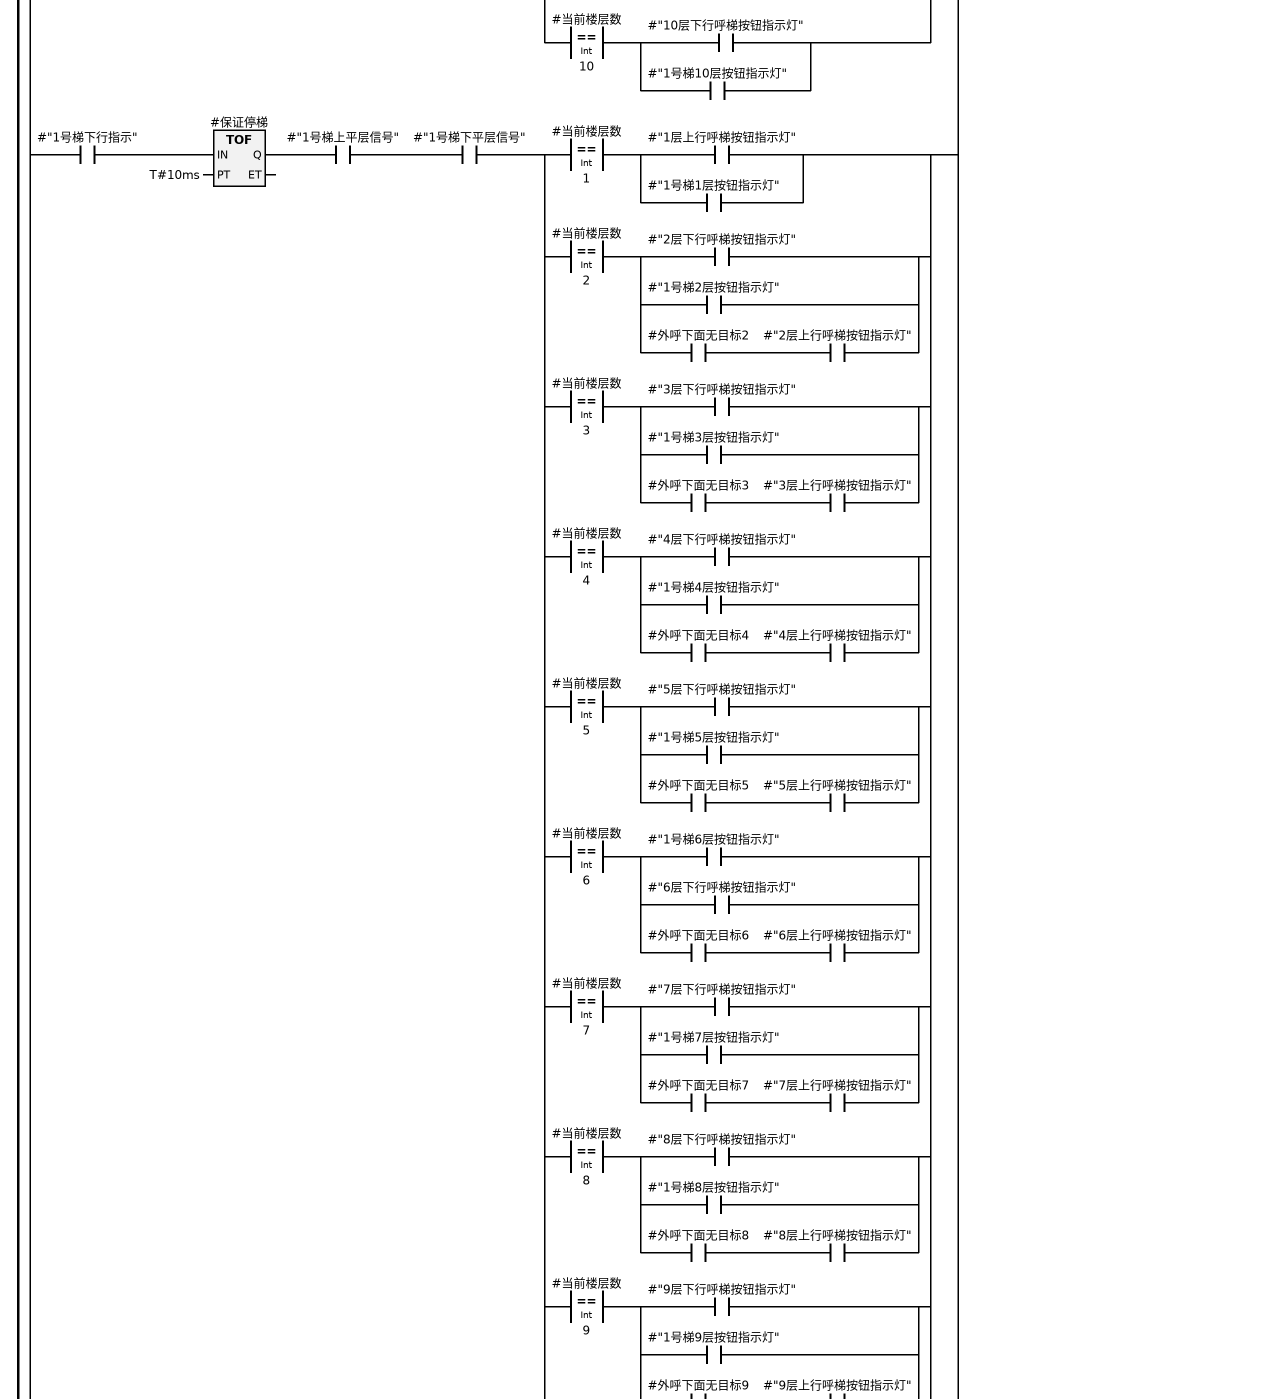
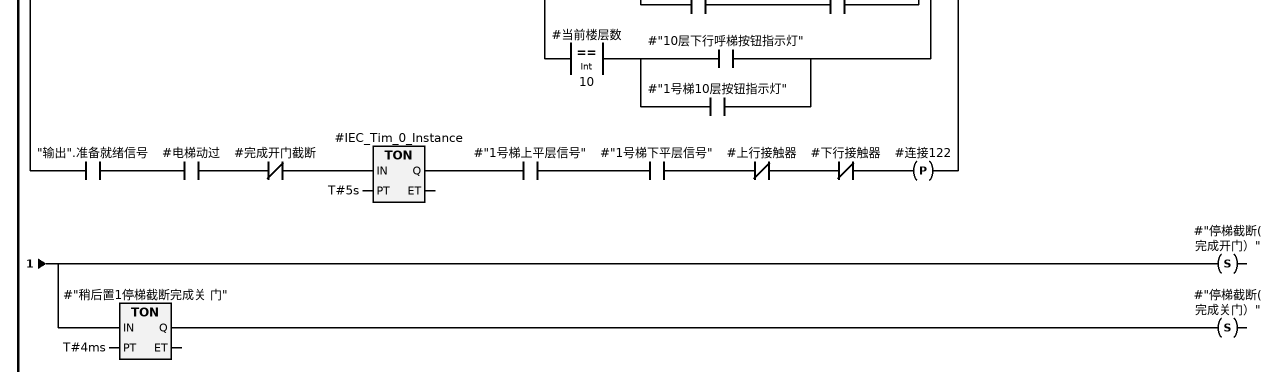
   #保证停梯上(IN := #"1号梯上行指示", PT := T#10ms);   // TOF
   #保证停梯(IN := #"1号梯下行指示", PT := T#10ms);   // TOF
   #IEC_Tim_0_Instance(IN := "输出".准备就绪信号 AND #电梯动过 AND NOT #完成开门截断, PT := T#5s);   // TON
   #_w1 := #IEC_Tim_0_Instance.Q AND #"1号梯上平层信号" AND #"1号梯下平层信号" AND NOT #上行接触器 AND NOT #下行接触器;
   #_w2 := #_w1 AND NOT #连接122;   // rising edge
   #连接122 := #_w1;
   #_w3 := ((#保证停梯上.Q AND #"1号梯上平层信号" AND #"1号梯下平层信号" AND (((#当前楼层数 = 1) AND (#"1层上行呼梯按钮指示灯" OR #"1号梯1层按钮指示灯")) OR ((#当前楼层数 = 2) AND (#"2层上行呼梯按钮指示灯" OR #"1号梯2层按钮指示灯" OR (#外呼上面无目标2 AND #"2层下行呼梯按钮指示灯"))) OR ((#当前楼层数 = 3) AND (#"3层上行呼梯按钮指示灯" OR #"1号梯3层按钮指示灯" OR (#外呼上面无目标3 AND #"3层下行呼梯按钮指示灯"))) OR ((#当前楼层数 = 4) AND (#"4层上行呼梯按钮指示灯" OR #"1号梯4层按钮指示灯" OR (#外呼上面无目标4 AND #"4层下行呼梯按钮指示灯"))) OR ((#当前楼层数 = 5) AND (#"5层上行呼梯按钮指示灯" OR #"1号梯5层按钮指示灯" OR (#外呼上面无目标5 AND #"5层下行呼梯按钮指示灯"))) OR ((#当前楼层数 = 6) AND (#"6层上行呼梯按钮指示灯" OR #"1号梯6层按钮指示灯" OR (#外呼上面无目标6 AND #"6层下行呼梯按钮指示灯"))) OR ((#当前楼层数 = 7) AND (#"7层上行呼梯按钮指示灯" OR #"1号梯7层按钮指示灯" OR (#外呼上面无目标7 AND #"7层下行呼梯按钮指示灯"))) OR ((#当前楼层数 = 8) AND (#"8层上行呼梯按钮指示灯" OR #"1号梯8层按钮指示灯" OR (#外呼上面无目标8 AND #"8层下行呼梯按钮指示灯"))) OR ((#当前楼层数 = 9) AND (#"9层上行呼梯按钮指示灯" OR #"1号梯9层按钮指示灯" OR (#外呼上面无目标9 AND #"9层下行呼梯按钮指示灯"))) OR ((#当前楼层数 = 10) AND (#"10层下行呼梯按钮指示灯" OR #"1号梯10层按钮指示灯")))) OR (#保证停梯.Q AND #"1号梯上平层信号" AND #"1号梯下平层信号" AND (((#当前楼层数 = 1) AND (#"1层上行呼梯按钮指示灯" OR #"1号梯1层按钮指示灯")) OR ((#当前楼层数 = 2) AND (#"2层下行呼梯按钮指示灯" OR #"1号梯2层按钮指示灯" OR (#外呼下面无目标2 AND #"2层上行呼梯按钮指示灯"))) OR ((#当前楼层数 = 3) AND (#"3层下行呼梯按钮指示灯" OR #"1号梯3层按钮指示灯" OR (#外呼下面无目标3 AND #"3层上行呼梯按钮指示灯"))) OR ((#当前楼层数 = 4) AND (#"4层下行呼梯按钮指示灯" OR #"1号梯4层按钮指示灯" OR (#外呼下面无目标4 AND #"4层上行呼梯按钮指示灯"))) OR ((#当前楼层数 = 5) AND (#"5层下行呼梯按钮指示灯" OR #"1号梯5层按钮指示灯" OR (#外呼下面无目标5 AND #"5层上行呼梯按钮指示灯"))) OR ((#当前楼层数 = 6) AND (#"1号梯6层按钮指示灯" OR #"6层下行呼梯按钮指示灯" OR (#外呼下面无目标6 AND #"6层上行呼梯按钮指示灯"))) OR ((#当前楼层数 = 7) AND (#"7层下行呼梯按钮指示灯" OR #"1号梯7层按钮指示灯" OR (#外呼下面无目标7 AND #"7层上行呼梯按钮指示灯"))) OR ((#当前楼层数 = 8) AND (#"8层下行呼梯按钮指示灯" OR #"1号梯8层按钮指示灯" OR (#外呼下面无目标8 AND #"8层上行呼梯按钮指示灯"))) OR ((#当前楼层数 = 9) AND (#"9层下行呼梯按钮指示灯" OR #"1号梯9层按钮指示灯" OR (#外呼下面无目标9 AND #"9层上行呼梯按钮指示灯"))) OR ((#当前楼层数 = 10) AND (#"10层下行呼梯按钮指示灯" OR #"1号梯10层按钮指示灯")))) OR #_w2) AND NOT #"1号梯检修信号" AND NOT #开门次数达到上限;
   IF #_w3 THEN #"停梯截断(完成开门）" := TRUE; END_IF;
   #"稍后置1停梯截断完成关 门"(IN := #_w3, PT := T#4ms);   // TON
   IF #"稍后置1停梯截断完成关 门".Q THEN #"停梯截断(完成关门）" := TRUE; END_IF;
END_REGION

REGION Network 2: 停梯后自主 开门
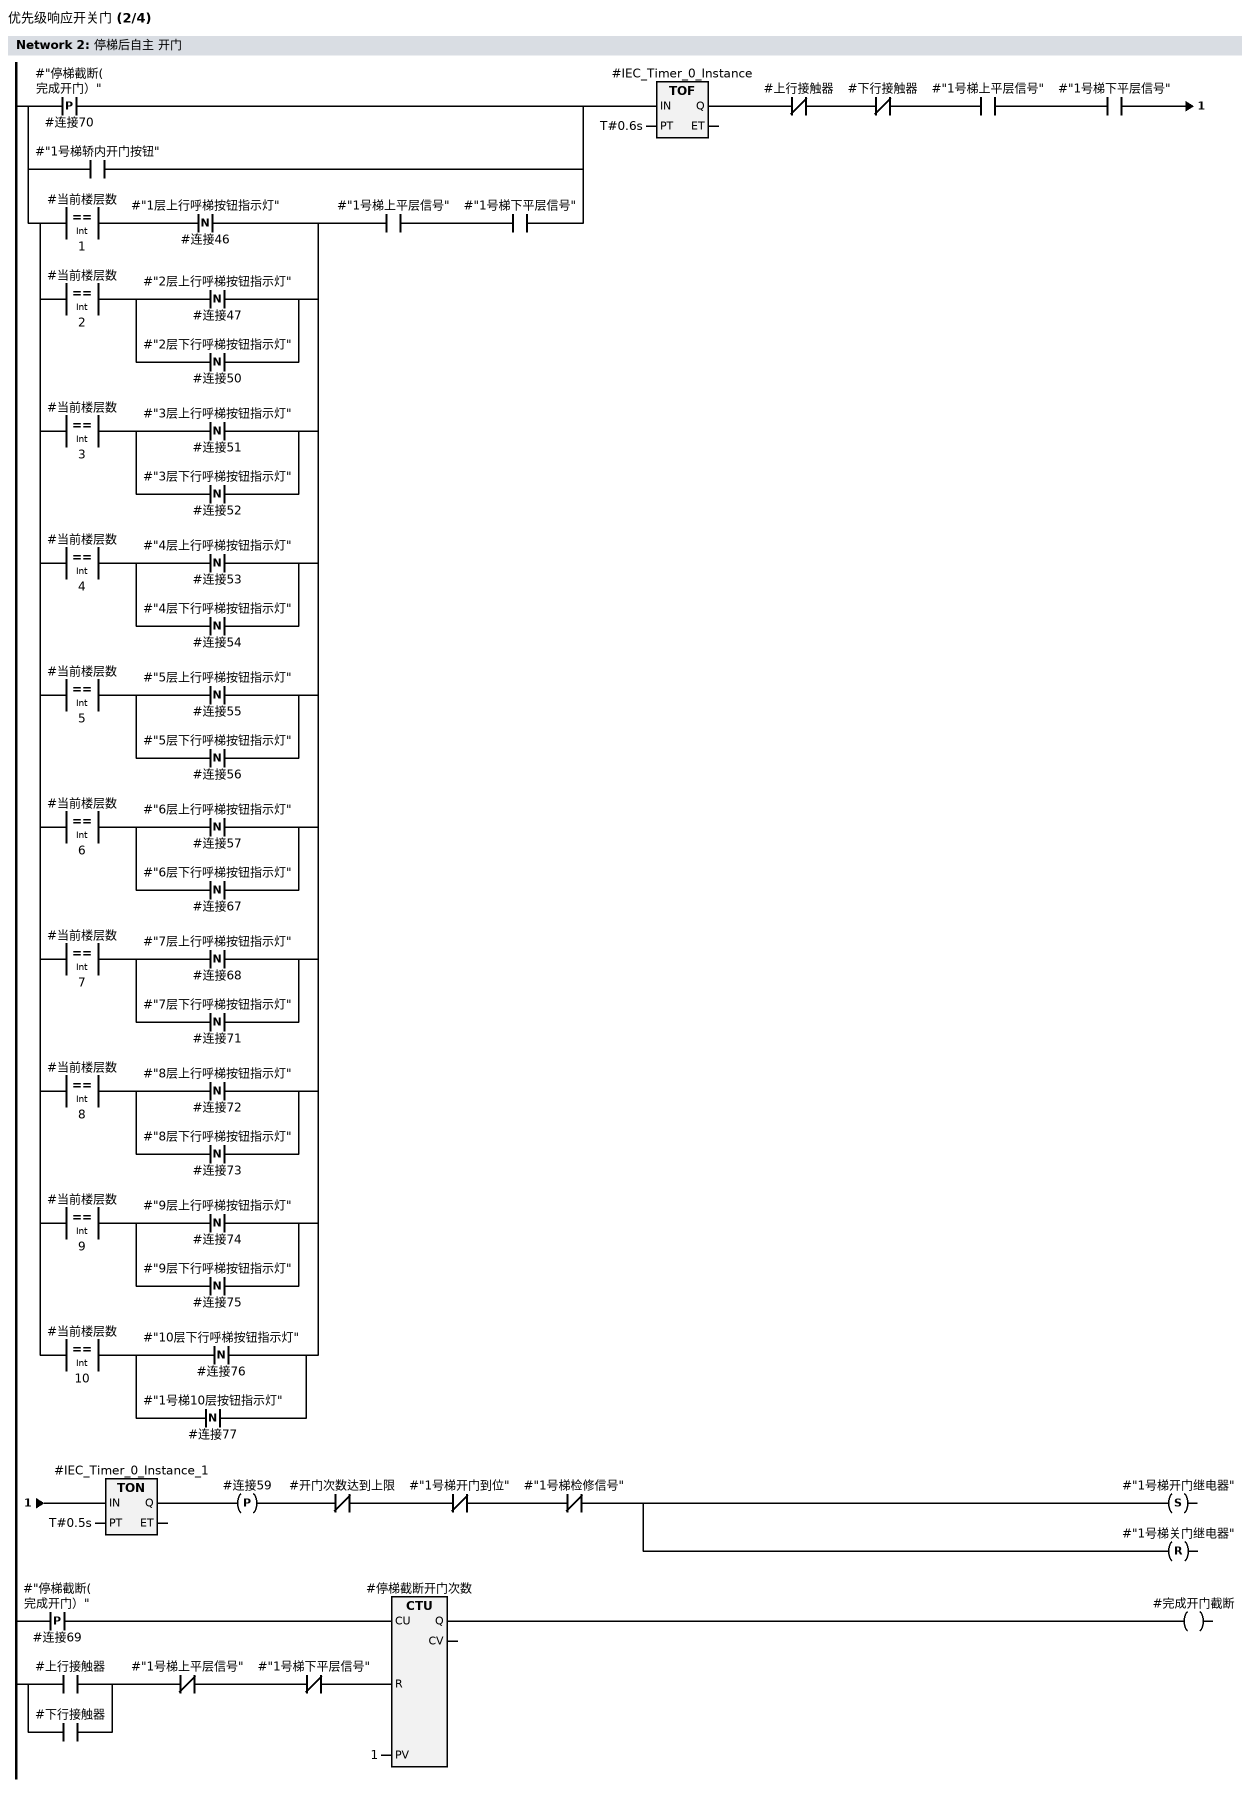
   #_w1 := #"停梯截断(完成开门）" AND NOT #连接70;   // rising edge of #"停梯截断(完成开门）"
   #连接70 := #"停梯截断(完成开门）";
   #_w2 := (#当前楼层数 = 1) AND NOT #"1层上行呼梯按钮指示灯" AND #连接46;   // falling edge of #"1层上行呼梯按钮指示灯"
   #连接46 := #"1层上行呼梯按钮指示灯";
   #_w3 := (#当前楼层数 = 2) AND NOT #"2层上行呼梯按钮指示灯" AND #连接47;   // falling edge of #"2层上行呼梯按钮指示灯"
   #连接47 := #"2层上行呼梯按钮指示灯";
   #_w4 := (#当前楼层数 = 2) AND NOT #"2层下行呼梯按钮指示灯" AND #连接50;   // falling edge of #"2层下行呼梯按钮指示灯"
   #连接50 := #"2层下行呼梯按钮指示灯";
   #_w5 := (#当前楼层数 = 3) AND NOT #"3层上行呼梯按钮指示灯" AND #连接51;   // falling edge of #"3层上行呼梯按钮指示灯"
   #连接51 := #"3层上行呼梯按钮指示灯";
   #_w6 := (#当前楼层数 = 3) AND NOT #"3层下行呼梯按钮指示灯" AND #连接52;   // falling edge of #"3层下行呼梯按钮指示灯"
   #连接52 := #"3层下行呼梯按钮指示灯";
   #_w7 := (#当前楼层数 = 4) AND NOT #"4层上行呼梯按钮指示灯" AND #连接53;   // falling edge of #"4层上行呼梯按钮指示灯"
   #连接53 := #"4层上行呼梯按钮指示灯";
   #_w8 := (#当前楼层数 = 4) AND NOT #"4层下行呼梯按钮指示灯" AND #连接54;   // falling edge of #"4层下行呼梯按钮指示灯"
   #连接54 := #"4层下行呼梯按钮指示灯";
   #_w9 := (#当前楼层数 = 5) AND NOT #"5层上行呼梯按钮指示灯" AND #连接55;   // falling edge of #"5层上行呼梯按钮指示灯"
   #连接55 := #"5层上行呼梯按钮指示灯";
   #_w10 := (#当前楼层数 = 5) AND NOT #"5层下行呼梯按钮指示灯" AND #连接56;   // falling edge of #"5层下行呼梯按钮指示灯"
   #连接56 := #"5层下行呼梯按钮指示灯";
   #_w11 := (#当前楼层数 = 6) AND NOT #"6层上行呼梯按钮指示灯" AND #连接57;   // falling edge of #"6层上行呼梯按钮指示灯"
   #连接57 := #"6层上行呼梯按钮指示灯";
   #_w12 := (#当前楼层数 = 6) AND NOT #"6层下行呼梯按钮指示灯" AND #连接67;   // falling edge of #"6层下行呼梯按钮指示灯"
   #连接67 := #"6层下行呼梯按钮指示灯";
   #_w13 := (#当前楼层数 = 7) AND NOT #"7层上行呼梯按钮指示灯" AND #连接68;   // falling edge of #"7层上行呼梯按钮指示灯"
   #连接68 := #"7层上行呼梯按钮指示灯";
   #_w14 := (#当前楼层数 = 7) AND NOT #"7层下行呼梯按钮指示灯" AND #连接71;   // falling edge of #"7层下行呼梯按钮指示灯"
   #连接71 := #"7层下行呼梯按钮指示灯";
   #_w15 := (#当前楼层数 = 8) AND NOT #"8层上行呼梯按钮指示灯" AND #连接72;   // falling edge of #"8层上行呼梯按钮指示灯"
   #连接72 := #"8层上行呼梯按钮指示灯";
   #_w16 := (#当前楼层数 = 8) AND NOT #"8层下行呼梯按钮指示灯" AND #连接73;   // falling edge of #"8层下行呼梯按钮指示灯"
   #连接73 := #"8层下行呼梯按钮指示灯";
   #_w17 := (#当前楼层数 = 9) AND NOT #"9层上行呼梯按钮指示灯" AND #连接74;   // falling edge of #"9层上行呼梯按钮指示灯"
   #连接74 := #"9层上行呼梯按钮指示灯";
   #_w18 := (#当前楼层数 = 9) AND NOT #"9层下行呼梯按钮指示灯" AND #连接75;   // falling edge of #"9层下行呼梯按钮指示灯"
   #连接75 := #"9层下行呼梯按钮指示灯";
   #_w19 := (#当前楼层数 = 10) AND NOT #"10层下行呼梯按钮指示灯" AND #连接76;   // falling edge of #"10层下行呼梯按钮指示灯"
   #连接76 := #"10层下行呼梯按钮指示灯";
   #_w20 := (#当前楼层数 = 10) AND NOT #"1号梯10层按钮指示灯" AND #连接77;   // falling edge of #"1号梯10层按钮指示灯"
   #连接77 := #"1号梯10层按钮指示灯";
   #IEC_Timer_0_Instance(IN := #_w1 OR #"1号梯轿内开门按钮" OR ((#_w2 OR #_w3 OR #_w4 OR #_w5 OR #_w6 OR #_w7 OR #_w8 OR #_w9 OR #_w10 OR #_w11 OR #_w12 OR #_w13 OR #_w14 OR #_w15 OR #_w16 OR #_w17 OR #_w18 OR #_w19 OR #_w20) AND #"1号梯上平层信号" AND #"1号梯下平层信号"),   // TOF
                         PT := T#0.6s);
   #IEC_Timer_0_Instance_1(IN := #IEC_Timer_0_Instance.Q AND NOT #上行接触器 AND NOT #下行接触器 AND #"1号梯上平层信号" AND #"1号梯下平层信号",   // TON
                           PT := T#0.5s);
   #_w21 := #IEC_Timer_0_Instance_1.Q AND NOT #连接59;   // rising edge
   #连接59 := #IEC_Timer_0_Instance_1.Q;
   IF #_w21 AND NOT #开门次数达到上限 AND NOT #"1号梯开门到位" AND NOT #"1号梯检修信号" THEN
       #"1号梯开门继电器" := TRUE;
       #"1号梯关门继电器" := FALSE;
   END_IF;
   #_w22 := #"停梯截断(完成开门）" AND NOT #连接69;   // rising edge of #"停梯截断(完成开门）"
   #连接69 := #"停梯截断(完成开门）";
   #停梯截断开门次数(CU := #_w22, R := (#上行接触器 OR #下行接触器) AND NOT #"1号梯上平层信号" AND NOT #"1号梯下平层信号", PV := 1);   // CTU
   #完成开门截断 := #停梯截断开门次数.Q;
END_REGION

REGION Network 3: 电梯自主完成开门关门
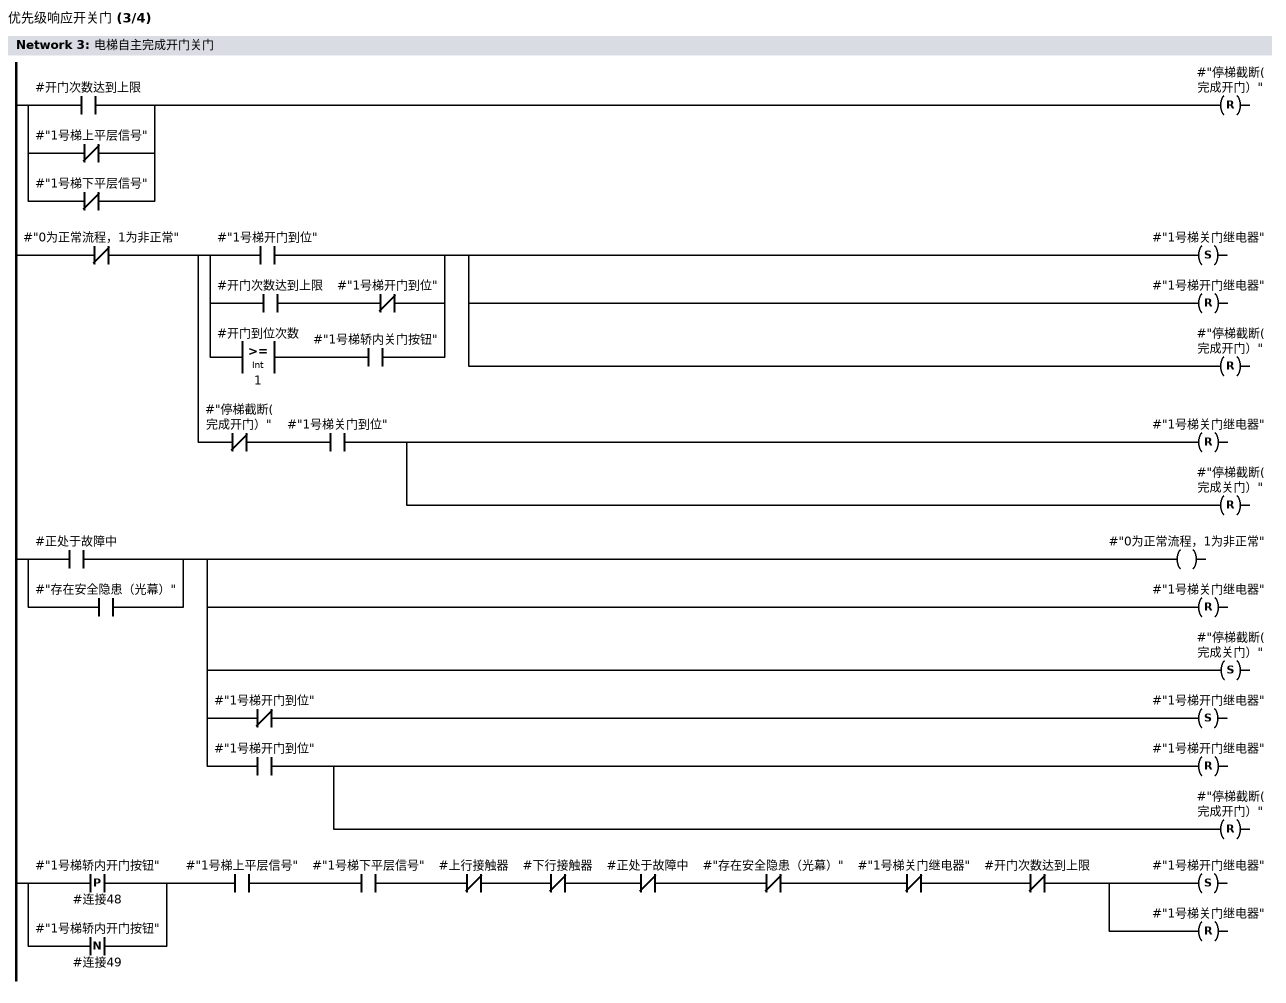
   RUNG wire#powerrail
      Contact( #开门次数达到上限 )
      wire#w1
      R_Coil( #"停梯截断(完成开门）" )
   END_RUNG
   RUNG wire#powerrail
      I_Contact( #"1号梯上平层信号" )
   END_RUNG wire#w1
   RUNG wire#powerrail
      I_Contact( #"1号梯下平层信号" )
   END_RUNG wire#w1
   RUNG wire#powerrail
      I_Contact( #"0为正常流程，1为非正常" )
      wire#w2
      Contact( #"1号梯开门到位" )
      wire#w3
      S_Coil( #"1号梯关门继电器" )
   END_RUNG
   RUNG wire#w2
      Contact( #开门次数达到上限 )
      I_Contact( #"1号梯开门到位" )
   END_RUNG wire#w3
   RUNG wire#w2
      { S7_Templates := "SrcType := Int" } GE_Contact(in1 := #开门到位次数, in2 := 1)
      Contact( #"1号梯轿内关门按钮" )
   END_RUNG wire#w3
   RUNG wire#w3
      R_Coil( #"1号梯开门继电器" )
   END_RUNG
   RUNG wire#w3
      R_Coil( #"停梯截断(完成开门）" )
   END_RUNG
   RUNG wire#w2
      I_Contact( #"停梯截断(完成开门）" )
      Contact( #"1号梯关门到位" )
      wire#w4
      R_Coil( #"1号梯关门继电器" )
   END_RUNG
   RUNG wire#w4
      R_Coil( #"停梯截断(完成关门）" )
   END_RUNG
   RUNG wire#powerrail
      Contact( #正处于故障中 )
      wire#w5
      Coil( #"0为正常流程，1为非正常" )
   END_RUNG
   RUNG wire#powerrail
      Contact( #"存在安全隐患（光幕）" )
   END_RUNG wire#w5
   RUNG wire#w5
      R_Coil( #"1号梯关门继电器" )
   END_RUNG
   RUNG wire#w5
      S_Coil( #"停梯截断(完成关门）" )
   END_RUNG
   RUNG wire#w5
      I_Contact( #"1号梯开门到位" )
      S_Coil( #"1号梯开门继电器" )
   END_RUNG
   RUNG wire#w5
      Contact( #"1号梯开门到位" )
      wire#w6
      R_Coil( #"1号梯开门继电器" )
   END_RUNG
   RUNG wire#w6
      R_Coil( #"停梯截断(完成开门）" )
   END_RUNG
   RUNG wire#powerrail
      P_Contact(operand := #"1号梯轿内开门按钮", bit := #连接48)
      wire#w7
      Contact( #"1号梯上平层信号" )
      Contact( #"1号梯下平层信号" )
      I_Contact( #上行接触器 )
      I_Contact( #下行接触器 )
      I_Contact( #正处于故障中 )
      I_Contact( #"存在安全隐患（光幕）" )
      I_Contact( #"1号梯关门继电器" )
      I_Contact( #开门次数达到上限 )
      wire#w8
      S_Coil( #"1号梯开门继电器" )
   END_RUNG
   RUNG wire#powerrail
      N_Contact(operand := #"1号梯轿内开门按钮", bit := #连接49)
   END_RUNG wire#w7
   RUNG wire#w8
      R_Coil( #"1号梯关门继电器" )
   END_RUNG
   // the same network as SCL:
   IF #开门次数达到上限 OR NOT #"1号梯上平层信号" OR NOT #"1号梯下平层信号" THEN #"停梯截断(完成开门）" := FALSE; END_IF;
   IF NOT #"0为正常流程，1为非正常" AND (#"1号梯开门到位" OR (#开门次数达到上限 AND NOT #"1号梯开门到位") OR ((#开门到位次数 >= 1) AND #"1号梯轿内关门按钮")) THEN
       #"1号梯关门继电器" := TRUE;
       #"1号梯开门继电器" := FALSE;
       #"停梯截断(完成开门）" := FALSE;
   END_IF;
   IF NOT #"0为正常流程，1为非正常" AND NOT #"停梯截断(完成开门）" AND #"1号梯关门到位" THEN
       #"1号梯关门继电器" := FALSE;
       #"停梯截断(完成关门）" := FALSE;
   END_IF;
   #"0为正常流程，1为非正常" := #正处于故障中 OR #"存在安全隐患（光幕）";
   IF #"0为正常流程，1为非正常" THEN
       #"1号梯关门继电器" := FALSE;
       #"停梯截断(完成关门）" := TRUE;
   END_IF;
   IF #"0为正常流程，1为非正常" AND NOT #"1号梯开门到位" THEN #"1号梯开门继电器" := TRUE; END_IF;
   IF #"0为正常流程，1为非正常" AND #"1号梯开门到位" THEN
       #"1号梯开门继电器" := FALSE;
       #"停梯截断(完成开门）" := FALSE;
   END_IF;
   #_w1 := #"1号梯轿内开门按钮" AND NOT #连接48;   // rising edge of #"1号梯轿内开门按钮"
   #连接48 := #"1号梯轿内开门按钮";
   #_w2 := NOT #"1号梯轿内开门按钮" AND #连接49;   // falling edge of #"1号梯轿内开门按钮"
   #连接49 := #"1号梯轿内开门按钮";
   IF (#_w1 OR #_w2) AND #"1号梯上平层信号" AND #"1号梯下平层信号" AND NOT #上行接触器 AND NOT #下行接触器 AND NOT #正处于故障中 AND NOT #"存在安全隐患（光幕）" AND NOT #"1号梯关门继电器" AND NOT #开门次数达到上限 THEN
       #"1号梯开门继电器" := TRUE;
       #"1号梯关门继电器" := FALSE;
   END_IF;
END_REGION

REGION Network 4: 检修与死机
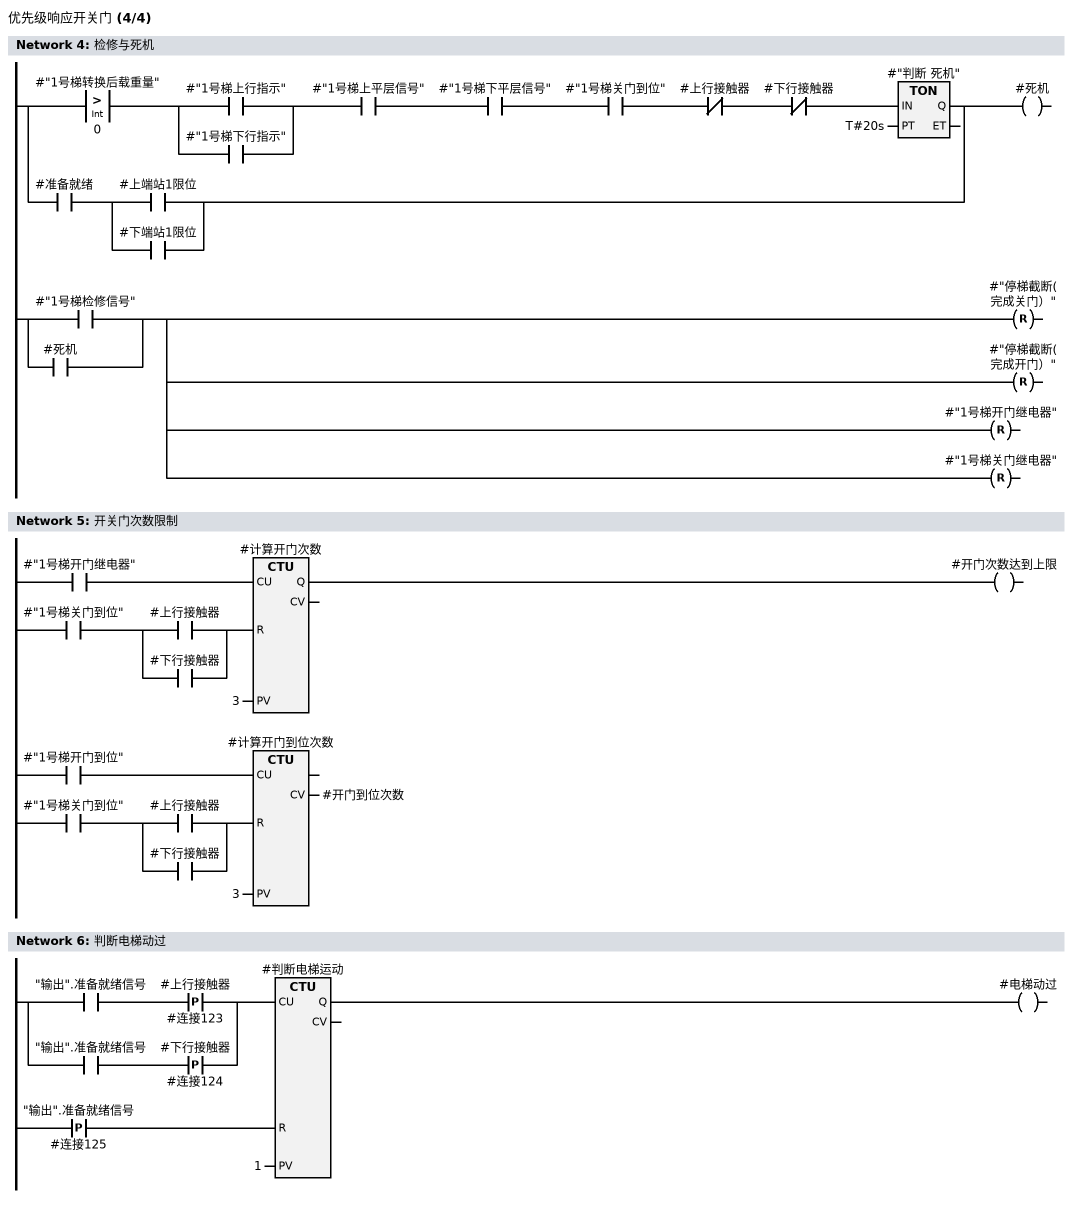
   #"判断 死机"(IN := (#"1号梯转换后载重量" > 0) AND (#"1号梯上行指示" OR #"1号梯下行指示") AND #"1号梯上平层信号" AND #"1号梯下平层信号" AND #"1号梯关门到位" AND NOT #上行接触器 AND NOT #下行接触器,   // TON
            PT := T#20s);
   #死机 := #"判断 死机".Q OR (#准备就绪 AND (#上端站1限位 OR #下端站1限位));
   IF #"1号梯检修信号" OR #死机 THEN
       #"停梯截断(完成关门）" := FALSE;
       #"停梯截断(完成开门）" := FALSE;
       #"1号梯开门继电器" := FALSE;
       #"1号梯关门继电器" := FALSE;
   END_IF;
END_REGION

REGION Network 5: 开关门次数限制
   #计算开门次数(CU := #"1号梯开门继电器", R := #"1号梯关门到位" AND (#上行接触器 OR #下行接触器), PV := 3);   // CTU
   #开门次数达到上限 := #计算开门次数.Q;
   #计算开门到位次数(CU := #"1号梯开门到位", R := #"1号梯关门到位" AND (#上行接触器 OR #下行接触器), PV := 3, CV => #开门到位次数);   // CTU
END_REGION

REGION Network 6: 判断电梯动过
   #_w1 := "输出".准备就绪信号 AND #上行接触器 AND NOT #连接123;   // rising edge of #上行接触器
   #连接123 := #上行接触器;
   #_w2 := "输出".准备就绪信号 AND #下行接触器 AND NOT #连接124;   // rising edge of #下行接触器
   #连接124 := #下行接触器;
   #_w3 := "输出".准备就绪信号 AND NOT #连接125;   // rising edge of "输出".准备就绪信号
   #连接125 := "输出".准备就绪信号;
   #判断电梯运动(CU := #_w1 OR #_w2, R := #_w3, PV := 1);   // CTU
   #电梯动过 := #判断电梯运动.Q;
END_REGION
END_FUNCTION_BLOCK

FUNCTION_BLOCK "高低速转换"   // FB13, LAD
{ S7_Optimized_Access := 'TRUE' }
VERSION : 0.1
   VAR_INPUT
      准备就绪 : Bool;
      初始化低速运行 : Bool;
      当前楼层数 : Int;
      "1层上行呼梯按钮指示灯" : Bool;
      "2层上行呼梯按钮指示灯" : Bool;
      "3层上行呼梯按钮指示灯" : Bool;
      "4层上行呼梯按钮指示灯" : Bool;
      "5层上行呼梯按钮指示灯" : Bool;
      "6层上行呼梯按钮指示灯" : Bool;
      "7层上行呼梯按钮指示灯" : Bool;
      "8层上行呼梯按钮指示灯" : Bool;
      "9层上行呼梯按钮指示灯" : Bool;
      "2层下行呼梯按钮指示灯" : Bool;
      "3层下行呼梯按钮指示灯" : Bool;
      "4层下行呼梯按钮指示灯" : Bool;
      "5层下行呼梯按钮指示灯" : Bool;
      "6层下行呼梯按钮指示灯" : Bool;
      "7层下行呼梯按钮指示灯" : Bool;
      "8层下行呼梯按钮指示灯" : Bool;
      "9层下行呼梯按钮指示灯" : Bool;
      "10层下行呼梯按钮指示灯" : Bool;
      "1号梯1层按钮指示灯" : Bool;
      "1号梯2层按钮指示灯" : Bool;
      "1号梯3层按钮指示灯" : Bool;
      "1号梯4层按钮指示灯" : Bool;
      "1号梯5层按钮指示灯" : Bool;
      "1号梯6层按钮指示灯" : Bool;
      "1号梯7层按钮指示灯" : Bool;
      "1号梯8层按钮指示灯" : Bool;
      "1号梯9层按钮指示灯" : Bool;
      "1号梯10层按钮指示灯" : Bool;
      正处于故障中 : Bool;
      "存在安全隐患（光幕）" : Bool;
      "1号梯上行指示" : Bool;
      "1号梯下行指示" : Bool;
      "1号梯检修信号" : Bool;
      "1号梯上行接触器" : Bool;
      "1号梯下行接触器" : Bool;
      "1号梯外呼上面无目标2" : Bool;
      "1号梯外呼上面无目标3" : Bool;
      "1号梯外呼上面无目标4" : Bool;
      "1号梯外呼上面无目标5" : Bool;
      "1号梯外呼上面无目标6" : Bool;
      "1号梯外呼上面无目标7" : Bool;
      "1号梯外呼上面无目标8" : Bool;
      "1号梯外呼上面无目标9" : Bool;
      "1号梯外呼下面无目标2" : Bool;
      "1号梯外呼下面无目标3" : Bool;
      "1号梯外呼下面无目标4" : Bool;
      "1号梯外呼下面无目标5" : Bool;
      "1号梯外呼下面无目标6" : Bool;
      "1号梯外呼下面无目标7" : Bool;
      "1号梯外呼下面无目标8" : Bool;
      "1号梯外呼下面无目标9" : Bool;
      初始化高速运行 : Bool;
   END_VAR
   VAR_OUTPUT
      "1号梯高速接触器" : Bool;
      "1号梯低速接触器" : Bool;
      将要停梯 : Bool;
   END_VAR
   VAR
      中间1 : Bool;
      中间2 : Bool;
      中间3 : Bool;
      中间4 : Bool;
      中间5 : Bool;
   END_VAR
BEGIN

REGION Network 1: 低速上下行（前正常指令，后最后指令）
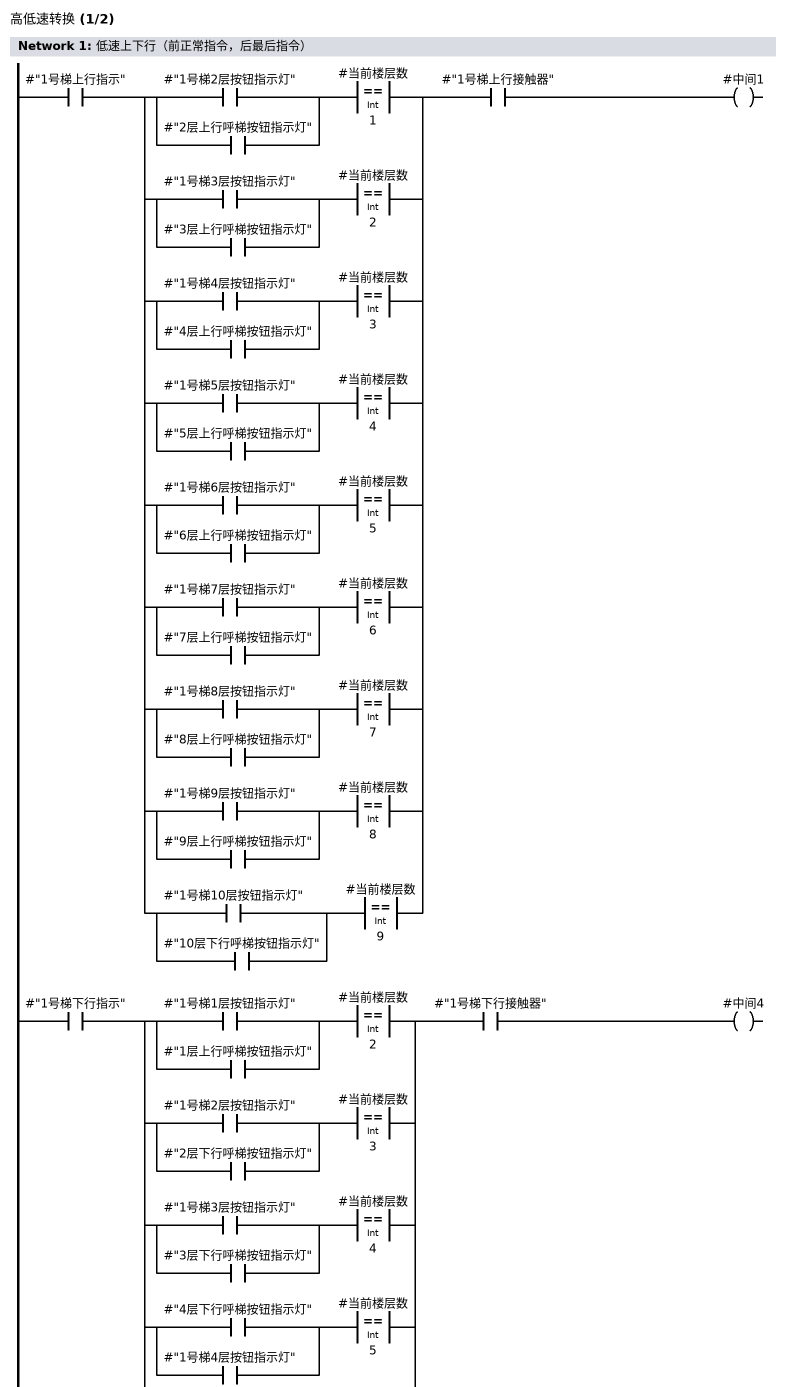
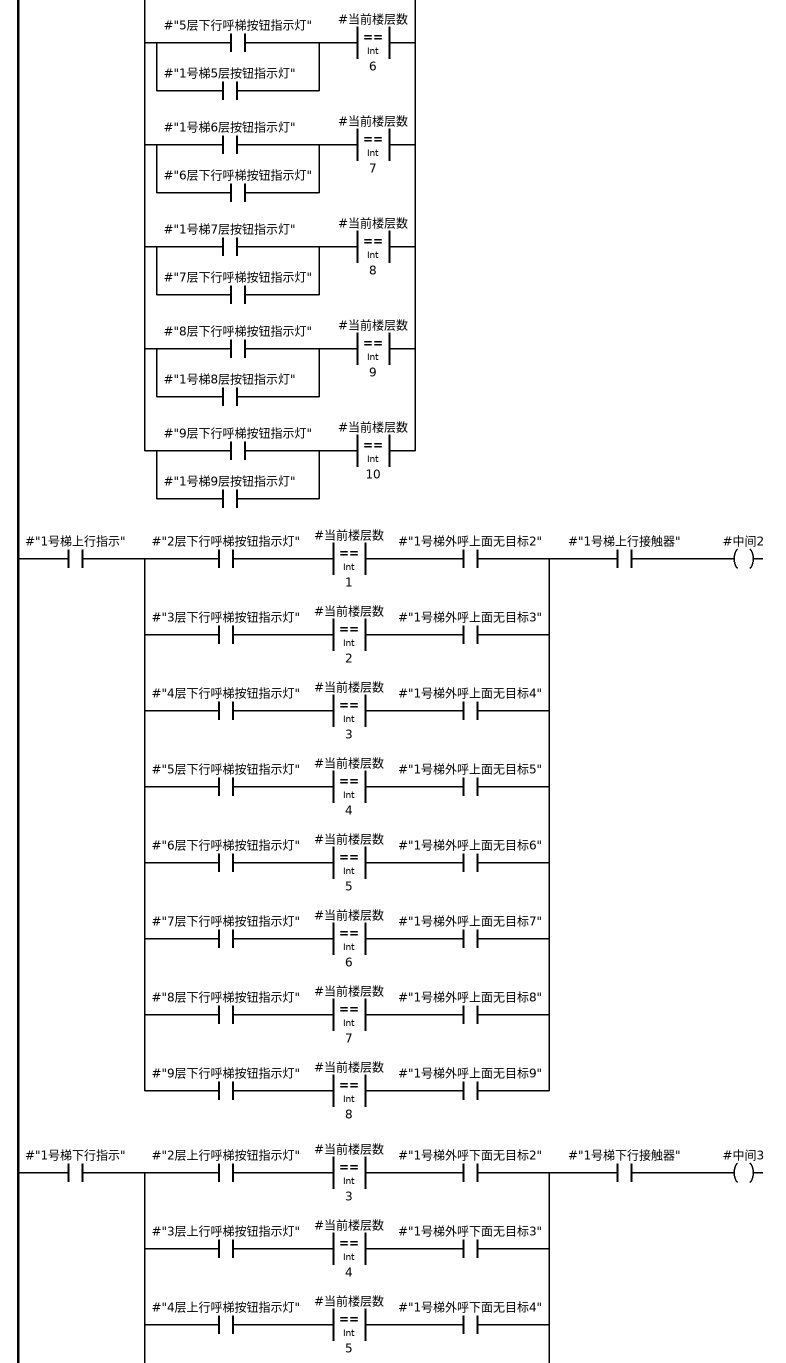
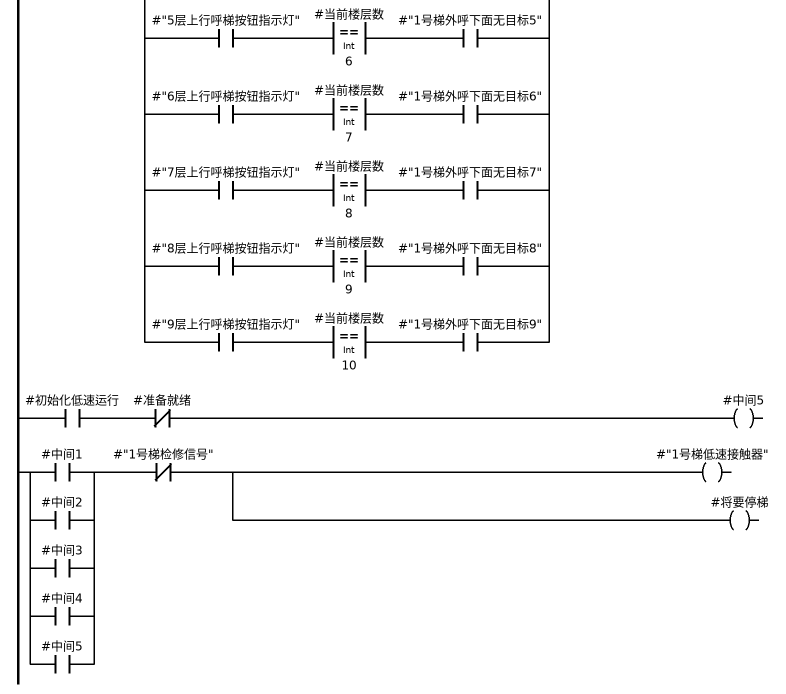
   RUNG wire#powerrail
      Contact( #"1号梯上行指示" )
      wire#w1
      Contact( #"1号梯2层按钮指示灯" )
      wire#w2
      { S7_Templates := "SrcType := Int" } EQ_Contact(in1 := #当前楼层数, in2 := 1)
      wire#w3
      Contact( #"1号梯上行接触器" )
      Coil( #中间1 )
   END_RUNG
   RUNG wire#w1
      Contact( #"2层上行呼梯按钮指示灯" )
   END_RUNG wire#w2
   RUNG wire#w1
      Contact( #"1号梯3层按钮指示灯" )
      wire#w4
      { S7_Templates := "SrcType := Int" } EQ_Contact(in1 := #当前楼层数, in2 := 2)
   END_RUNG wire#w3
   RUNG wire#w1
      Contact( #"3层上行呼梯按钮指示灯" )
   END_RUNG wire#w4
   RUNG wire#w1
      Contact( #"1号梯4层按钮指示灯" )
      wire#w5
      { S7_Templates := "SrcType := Int" } EQ_Contact(in1 := #当前楼层数, in2 := 3)
   END_RUNG wire#w3
   RUNG wire#w1
      Contact( #"4层上行呼梯按钮指示灯" )
   END_RUNG wire#w5
   RUNG wire#w1
      Contact( #"1号梯5层按钮指示灯" )
      wire#w6
      { S7_Templates := "SrcType := Int" } EQ_Contact(in1 := #当前楼层数, in2 := 4)
   END_RUNG wire#w3
   RUNG wire#w1
      Contact( #"5层上行呼梯按钮指示灯" )
   END_RUNG wire#w6
   RUNG wire#w1
      Contact( #"1号梯6层按钮指示灯" )
      wire#w7
      { S7_Templates := "SrcType := Int" } EQ_Contact(in1 := #当前楼层数, in2 := 5)
   END_RUNG wire#w3
   RUNG wire#w1
      Contact( #"6层上行呼梯按钮指示灯" )
   END_RUNG wire#w7
   RUNG wire#w1
      Contact( #"1号梯7层按钮指示灯" )
      wire#w8
      { S7_Templates := "SrcType := Int" } EQ_Contact(in1 := #当前楼层数, in2 := 6)
   END_RUNG wire#w3
   RUNG wire#w1
      Contact( #"7层上行呼梯按钮指示灯" )
   END_RUNG wire#w8
   RUNG wire#w1
      Contact( #"1号梯8层按钮指示灯" )
      wire#w9
      { S7_Templates := "SrcType := Int" } EQ_Contact(in1 := #当前楼层数, in2 := 7)
   END_RUNG wire#w3
   RUNG wire#w1
      Contact( #"8层上行呼梯按钮指示灯" )
   END_RUNG wire#w9
   RUNG wire#w1
      Contact( #"1号梯9层按钮指示灯" )
      wire#w10
      { S7_Templates := "SrcType := Int" } EQ_Contact(in1 := #当前楼层数, in2 := 8)
   END_RUNG wire#w3
   RUNG wire#w1
      Contact( #"9层上行呼梯按钮指示灯" )
   END_RUNG wire#w10
   RUNG wire#w1
      Contact( #"1号梯10层按钮指示灯" )
      wire#w11
      { S7_Templates := "SrcType := Int" } EQ_Contact(in1 := #当前楼层数, in2 := 9)
   END_RUNG wire#w3
   RUNG wire#w1
      Contact( #"10层下行呼梯按钮指示灯" )
   END_RUNG wire#w11
   RUNG wire#powerrail
      Contact( #"1号梯下行指示" )
      wire#w12
      Contact( #"1号梯1层按钮指示灯" )
      wire#w13
      { S7_Templates := "SrcType := Int" } EQ_Contact(in1 := #当前楼层数, in2 := 2)
      wire#w14
      Contact( #"1号梯下行接触器" )
      Coil( #中间4 )
   END_RUNG
   RUNG wire#w12
      Contact( #"1层上行呼梯按钮指示灯" )
   END_RUNG wire#w13
   RUNG wire#w12
      Contact( #"1号梯2层按钮指示灯" )
      wire#w15
      { S7_Templates := "SrcType := Int" } EQ_Contact(in1 := #当前楼层数, in2 := 3)
   END_RUNG wire#w14
   RUNG wire#w12
      Contact( #"2层下行呼梯按钮指示灯" )
   END_RUNG wire#w15
   RUNG wire#w12
      Contact( #"1号梯3层按钮指示灯" )
      wire#w16
      { S7_Templates := "SrcType := Int" } EQ_Contact(in1 := #当前楼层数, in2 := 4)
   END_RUNG wire#w14
   RUNG wire#w12
      Contact( #"3层下行呼梯按钮指示灯" )
   END_RUNG wire#w16
   RUNG wire#w12
      Contact( #"4层下行呼梯按钮指示灯" )
      wire#w17
      { S7_Templates := "SrcType := Int" } EQ_Contact(in1 := #当前楼层数, in2 := 5)
   END_RUNG wire#w14
   RUNG wire#w12
      Contact( #"1号梯4层按钮指示灯" )
   END_RUNG wire#w17
   RUNG wire#w12
      Contact( #"5层下行呼梯按钮指示灯" )
      wire#w18
      { S7_Templates := "SrcType := Int" } EQ_Contact(in1 := #当前楼层数, in2 := 6)
   END_RUNG wire#w14
   RUNG wire#w12
      Contact( #"1号梯5层按钮指示灯" )
   END_RUNG wire#w18
   RUNG wire#w12
      Contact( #"1号梯6层按钮指示灯" )
      wire#w19
      { S7_Templates := "SrcType := Int" } EQ_Contact(in1 := #当前楼层数, in2 := 7)
   END_RUNG wire#w14
   RUNG wire#w12
      Contact( #"6层下行呼梯按钮指示灯" )
   END_RUNG wire#w19
   RUNG wire#w12
      Contact( #"1号梯7层按钮指示灯" )
      wire#w20
      { S7_Templates := "SrcType := Int" } EQ_Contact(in1 := #当前楼层数, in2 := 8)
   END_RUNG wire#w14
   RUNG wire#w12
      Contact( #"7层下行呼梯按钮指示灯" )
   END_RUNG wire#w20
   RUNG wire#w12
      Contact( #"8层下行呼梯按钮指示灯" )
      wire#w21
      { S7_Templates := "SrcType := Int" } EQ_Contact(in1 := #当前楼层数, in2 := 9)
   END_RUNG wire#w14
   RUNG wire#w12
      Contact( #"1号梯8层按钮指示灯" )
   END_RUNG wire#w21
   RUNG wire#w12
      Contact( #"9层下行呼梯按钮指示灯" )
      wire#w22
      { S7_Templates := "SrcType := Int" } EQ_Contact(in1 := #当前楼层数, in2 := 10)
   END_RUNG wire#w14
   RUNG wire#w12
      Contact( #"1号梯9层按钮指示灯" )
   END_RUNG wire#w22
   RUNG wire#powerrail
      Contact( #"1号梯上行指示" )
      wire#w23
      Contact( #"2层下行呼梯按钮指示灯" )
      { S7_Templates := "SrcType := Int" } EQ_Contact(in1 := #当前楼层数, in2 := 1)
      Contact( #"1号梯外呼上面无目标2" )
      wire#w24
      Contact( #"1号梯上行接触器" )
      Coil( #中间2 )
   END_RUNG
   RUNG wire#w23
      Contact( #"3层下行呼梯按钮指示灯" )
      { S7_Templates := "SrcType := Int" } EQ_Contact(in1 := #当前楼层数, in2 := 2)
      Contact( #"1号梯外呼上面无目标3" )
   END_RUNG wire#w24
   RUNG wire#w23
      Contact( #"4层下行呼梯按钮指示灯" )
      { S7_Templates := "SrcType := Int" } EQ_Contact(in1 := #当前楼层数, in2 := 3)
      Contact( #"1号梯外呼上面无目标4" )
   END_RUNG wire#w24
   RUNG wire#w23
      Contact( #"5层下行呼梯按钮指示灯" )
      { S7_Templates := "SrcType := Int" } EQ_Contact(in1 := #当前楼层数, in2 := 4)
      Contact( #"1号梯外呼上面无目标5" )
   END_RUNG wire#w24
   RUNG wire#w23
      Contact( #"6层下行呼梯按钮指示灯" )
      { S7_Templates := "SrcType := Int" } EQ_Contact(in1 := #当前楼层数, in2 := 5)
      Contact( #"1号梯外呼上面无目标6" )
   END_RUNG wire#w24
   RUNG wire#w23
      Contact( #"7层下行呼梯按钮指示灯" )
      { S7_Templates := "SrcType := Int" } EQ_Contact(in1 := #当前楼层数, in2 := 6)
      Contact( #"1号梯外呼上面无目标7" )
   END_RUNG wire#w24
   RUNG wire#w23
      Contact( #"8层下行呼梯按钮指示灯" )
      { S7_Templates := "SrcType := Int" } EQ_Contact(in1 := #当前楼层数, in2 := 7)
      Contact( #"1号梯外呼上面无目标8" )
   END_RUNG wire#w24
   RUNG wire#w23
      Contact( #"9层下行呼梯按钮指示灯" )
      { S7_Templates := "SrcType := Int" } EQ_Contact(in1 := #当前楼层数, in2 := 8)
      Contact( #"1号梯外呼上面无目标9" )
   END_RUNG wire#w24
   RUNG wire#powerrail
      Contact( #"1号梯下行指示" )
      wire#w25
      Contact( #"2层上行呼梯按钮指示灯" )
      { S7_Templates := "SrcType := Int" } EQ_Contact(in1 := #当前楼层数, in2 := 3)
      Contact( #"1号梯外呼下面无目标2" )
      wire#w26
      Contact( #"1号梯下行接触器" )
      Coil( #中间3 )
   END_RUNG
   RUNG wire#w25
      Contact( #"3层上行呼梯按钮指示灯" )
      { S7_Templates := "SrcType := Int" } EQ_Contact(in1 := #当前楼层数, in2 := 4)
      Contact( #"1号梯外呼下面无目标3" )
   END_RUNG wire#w26
   RUNG wire#w25
      Contact( #"4层上行呼梯按钮指示灯" )
      { S7_Templates := "SrcType := Int" } EQ_Contact(in1 := #当前楼层数, in2 := 5)
      Contact( #"1号梯外呼下面无目标4" )
   END_RUNG wire#w26
   RUNG wire#w25
      Contact( #"5层上行呼梯按钮指示灯" )
      { S7_Templates := "SrcType := Int" } EQ_Contact(in1 := #当前楼层数, in2 := 6)
      Contact( #"1号梯外呼下面无目标5" )
   END_RUNG wire#w26
   RUNG wire#w25
      Contact( #"6层上行呼梯按钮指示灯" )
      { S7_Templates := "SrcType := Int" } EQ_Contact(in1 := #当前楼层数, in2 := 7)
      Contact( #"1号梯外呼下面无目标6" )
   END_RUNG wire#w26
   RUNG wire#w25
      Contact( #"7层上行呼梯按钮指示灯" )
      { S7_Templates := "SrcType := Int" } EQ_Contact(in1 := #当前楼层数, in2 := 8)
      Contact( #"1号梯外呼下面无目标7" )
   END_RUNG wire#w26
   RUNG wire#w25
      Contact( #"8层上行呼梯按钮指示灯" )
      { S7_Templates := "SrcType := Int" } EQ_Contact(in1 := #当前楼层数, in2 := 9)
      Contact( #"1号梯外呼下面无目标8" )
   END_RUNG wire#w26
   RUNG wire#w25
      Contact( #"9层上行呼梯按钮指示灯" )
      { S7_Templates := "SrcType := Int" } EQ_Contact(in1 := #当前楼层数, in2 := 10)
      Contact( #"1号梯外呼下面无目标9" )
   END_RUNG wire#w26
   RUNG wire#powerrail
      Contact( #初始化低速运行 )
      I_Contact( #准备就绪 )
      Coil( #中间5 )
   END_RUNG
   RUNG wire#powerrail
      Contact( #中间1 )
      wire#w27
      I_Contact( #"1号梯检修信号" )
      wire#w28
      Coil( #"1号梯低速接触器" )
   END_RUNG
   RUNG wire#powerrail
      Contact( #中间2 )
   END_RUNG wire#w27
   RUNG wire#powerrail
      Contact( #中间3 )
   END_RUNG wire#w27
   RUNG wire#powerrail
      Contact( #中间4 )
   END_RUNG wire#w27
   RUNG wire#powerrail
      Contact( #中间5 )
   END_RUNG wire#w27
   RUNG wire#w28
      Coil( #将要停梯 )
   END_RUNG
   // the same network as SCL:
   #中间1 := #"1号梯上行指示" AND (((#"1号梯2层按钮指示灯" OR #"2层上行呼梯按钮指示灯") AND (#当前楼层数 = 1)) OR ((#"1号梯3层按钮指示灯" OR #"3层上行呼梯按钮指示灯") AND (#当前楼层数 = 2)) OR ((#"1号梯4层按钮指示灯" OR #"4层上行呼梯按钮指示灯") AND (#当前楼层数 = 3)) OR ((#"1号梯5层按钮指示灯" OR #"5层上行呼梯按钮指示灯") AND (#当前楼层数 = 4)) OR ((#"1号梯6层按钮指示灯" OR #"6层上行呼梯按钮指示灯") AND (#当前楼层数 = 5)) OR ((#"1号梯7层按钮指示灯" OR #"7层上行呼梯按钮指示灯") AND (#当前楼层数 = 6)) OR ((#"1号梯8层按钮指示灯" OR #"8层上行呼梯按钮指示灯") AND (#当前楼层数 = 7)) OR ((#"1号梯9层按钮指示灯" OR #"9层上行呼梯按钮指示灯") AND (#当前楼层数 = 8)) OR ((#"1号梯10层按钮指示灯" OR #"10层下行呼梯按钮指示灯") AND (#当前楼层数 = 9))) AND #"1号梯上行接触器";
   #中间4 := #"1号梯下行指示" AND (((#"1号梯1层按钮指示灯" OR #"1层上行呼梯按钮指示灯") AND (#当前楼层数 = 2)) OR ((#"1号梯2层按钮指示灯" OR #"2层下行呼梯按钮指示灯") AND (#当前楼层数 = 3)) OR ((#"1号梯3层按钮指示灯" OR #"3层下行呼梯按钮指示灯") AND (#当前楼层数 = 4)) OR ((#"4层下行呼梯按钮指示灯" OR #"1号梯4层按钮指示灯") AND (#当前楼层数 = 5)) OR ((#"5层下行呼梯按钮指示灯" OR #"1号梯5层按钮指示灯") AND (#当前楼层数 = 6)) OR ((#"1号梯6层按钮指示灯" OR #"6层下行呼梯按钮指示灯") AND (#当前楼层数 = 7)) OR ((#"1号梯7层按钮指示灯" OR #"7层下行呼梯按钮指示灯") AND (#当前楼层数 = 8)) OR ((#"8层下行呼梯按钮指示灯" OR #"1号梯8层按钮指示灯") AND (#当前楼层数 = 9)) OR ((#"9层下行呼梯按钮指示灯" OR #"1号梯9层按钮指示灯") AND (#当前楼层数 = 10))) AND #"1号梯下行接触器";
   #中间2 := #"1号梯上行指示" AND ((#"2层下行呼梯按钮指示灯" AND (#当前楼层数 = 1) AND #"1号梯外呼上面无目标2") OR (#"3层下行呼梯按钮指示灯" AND (#当前楼层数 = 2) AND #"1号梯外呼上面无目标3") OR (#"4层下行呼梯按钮指示灯" AND (#当前楼层数 = 3) AND #"1号梯外呼上面无目标4") OR (#"5层下行呼梯按钮指示灯" AND (#当前楼层数 = 4) AND #"1号梯外呼上面无目标5") OR (#"6层下行呼梯按钮指示灯" AND (#当前楼层数 = 5) AND #"1号梯外呼上面无目标6") OR (#"7层下行呼梯按钮指示灯" AND (#当前楼层数 = 6) AND #"1号梯外呼上面无目标7") OR (#"8层下行呼梯按钮指示灯" AND (#当前楼层数 = 7) AND #"1号梯外呼上面无目标8") OR (#"9层下行呼梯按钮指示灯" AND (#当前楼层数 = 8) AND #"1号梯外呼上面无目标9")) AND #"1号梯上行接触器";
   #中间3 := #"1号梯下行指示" AND ((#"2层上行呼梯按钮指示灯" AND (#当前楼层数 = 3) AND #"1号梯外呼下面无目标2") OR (#"3层上行呼梯按钮指示灯" AND (#当前楼层数 = 4) AND #"1号梯外呼下面无目标3") OR (#"4层上行呼梯按钮指示灯" AND (#当前楼层数 = 5) AND #"1号梯外呼下面无目标4") OR (#"5层上行呼梯按钮指示灯" AND (#当前楼层数 = 6) AND #"1号梯外呼下面无目标5") OR (#"6层上行呼梯按钮指示灯" AND (#当前楼层数 = 7) AND #"1号梯外呼下面无目标6") OR (#"7层上行呼梯按钮指示灯" AND (#当前楼层数 = 8) AND #"1号梯外呼下面无目标7") OR (#"8层上行呼梯按钮指示灯" AND (#当前楼层数 = 9) AND #"1号梯外呼下面无目标8") OR (#"9层上行呼梯按钮指示灯" AND (#当前楼层数 = 10) AND #"1号梯外呼下面无目标9")) AND #"1号梯下行接触器";
   #中间5 := #初始化低速运行 AND NOT #准备就绪;
   #"1号梯低速接触器" := (#中间1 OR #中间2 OR #中间3 OR #中间4 OR #中间5) AND NOT #"1号梯检修信号";
   #将要停梯 := #"1号梯低速接触器";
END_REGION

REGION Network 2: 初始化高速
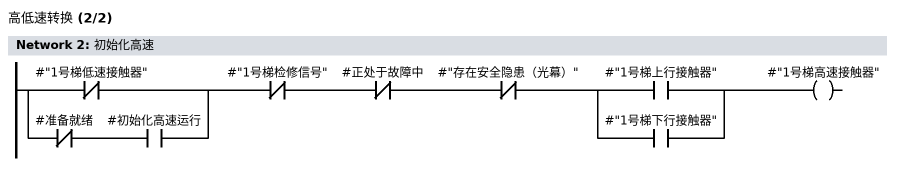
   RUNG wire#powerrail
      I_Contact( #"1号梯低速接触器" )
      wire#w1
      I_Contact( #"1号梯检修信号" )
      I_Contact( #正处于故障中 )
      I_Contact( #"存在安全隐患（光幕）" )
      wire#w2
      Contact( #"1号梯上行接触器" )
      wire#w3
      Coil( #"1号梯高速接触器" )
   END_RUNG
   RUNG wire#powerrail
      I_Contact( #准备就绪 )
      Contact( #初始化高速运行 )
   END_RUNG wire#w1
   RUNG wire#w2
      Contact( #"1号梯下行接触器" )
   END_RUNG wire#w3
   // the same network as SCL:
   #"1号梯高速接触器" := (NOT #"1号梯低速接触器" OR (NOT #准备就绪 AND #初始化高速运行)) AND NOT #"1号梯检修信号" AND NOT #正处于故障中 AND NOT #"存在安全隐患（光幕）" AND (#"1号梯上行接触器" OR #"1号梯下行接触器");
END_REGION
END_FUNCTION_BLOCK

FUNCTION_BLOCK "照明，风扇，数码管"   // FB15, LAD
{ S7_Optimized_Access := 'TRUE' }
VERSION : 0.1
   VAR_INPUT
      "1号梯光幕信号" : Bool;
      "1号梯开门到位" : Bool;
      "1号梯当前载重量" : Word;
      当前楼层数 : Int;
      "1号梯检修信号" : Bool;
      开门继电器 : Bool;
      关门继电器 : Bool;
      关门到位 : Bool;
      转换后载重量 : Int;
      载重限额 : Int;
      上行接触器 : Bool;
      下行接触器 : Bool;
   END_VAR
   VAR_OUTPUT
      正处于故障中 : Bool;
      安全隐患 : Bool;
      "1号梯LEDa" : Bool;
      "1号梯LEDb" : Bool;
      "1号梯LEDc" : Bool;
      "1号梯LEDd" : Bool;
      "1号梯LEDe" : Bool;
      "1号梯LEDf" : Bool;
      "1号梯LEDg" : Bool;
      "1号梯LEDh" : Bool;
      "1号梯LEDi" : Bool;
      "1号梯LEDj" : Bool;
      "1号梯LEDk" : Bool;
      "1号梯LEDl" : Bool;
      "1号梯LEDm" : Bool;
      "1号梯LEDn" : Bool;
      "1号梯照明指示" : Bool;
      "1号梯风扇指示" : Bool;
      "1号梯满载指示" : Bool;
      "1号梯故障指示" : Bool;
   END_VAR
   VAR
      开启故障闪烁 : Bool;
      停止故障闪烁 : Bool;
      连接99 : Bool;
      连接100 : Bool;
      连接104 : Bool;
      连接105 : Bool;
      连接106 : Bool;
      故障闪烁 : TON_TIME;
      "故障指示 闪烁" : TON_TIME;
      "IEC_Timer_ 0_Instance" : TON_TIME;
      IEC_Timer_0_Instance : TOF_TIME;
   END_VAR
   VAR_TEMP   // added for the SCL form of the ladder/FBD networks
      _w1 : Bool;
      _w2 : Bool;
      _w3 : Bool;
   END_VAR
BEGIN

REGION Network 1: 照明与风扇
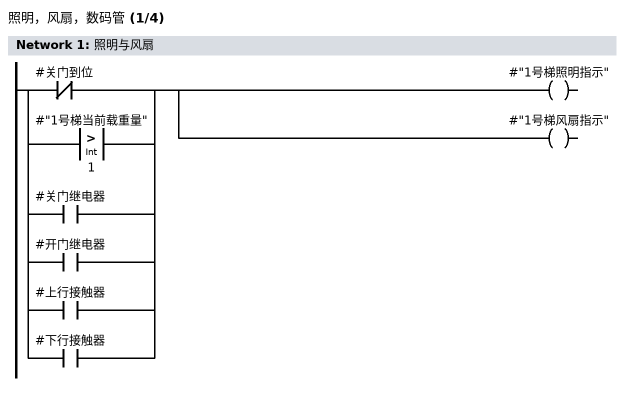
   RUNG wire#powerrail
      I_Contact( #关门到位 )
      wire#w1
      Coil( #"1号梯照明指示" )
   END_RUNG
   RUNG wire#powerrail
      { S7_Templates := "SrcType := Int" } GT_Contact(in1 := #"1号梯当前载重量", in2 := 1)
   END_RUNG wire#w1
   RUNG wire#powerrail
      Contact( #关门继电器 )
   END_RUNG wire#w1
   RUNG wire#powerrail
      Contact( #开门继电器 )
   END_RUNG wire#w1
   RUNG wire#powerrail
      Contact( #上行接触器 )
   END_RUNG wire#w1
   RUNG wire#powerrail
      Contact( #下行接触器 )
   END_RUNG wire#w1
   RUNG wire#w1
      Coil( #"1号梯风扇指示" )
   END_RUNG
   // the same network as SCL:
   #"1号梯照明指示" := NOT #关门到位 OR (#"1号梯当前载重量" > 1) OR #关门继电器 OR #开门继电器 OR #上行接触器 OR #下行接触器;
   #"1号梯风扇指示" := #"1号梯照明指示";
END_REGION

REGION Network 2: 数码管
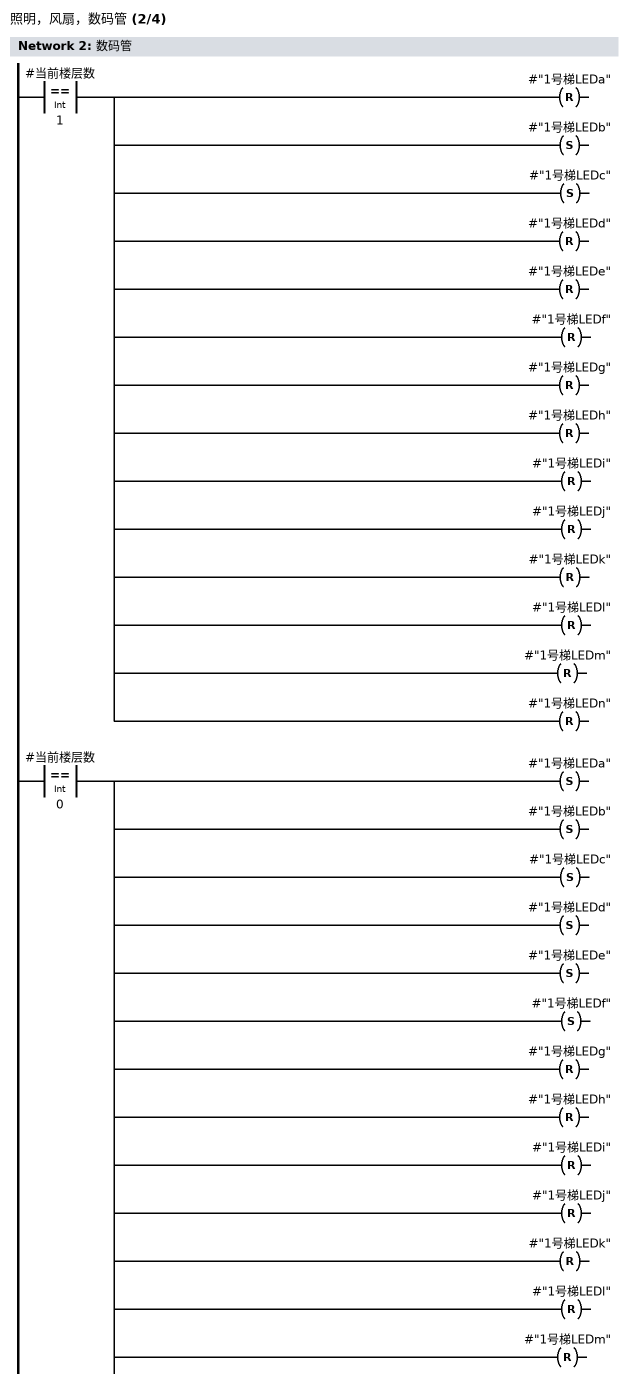
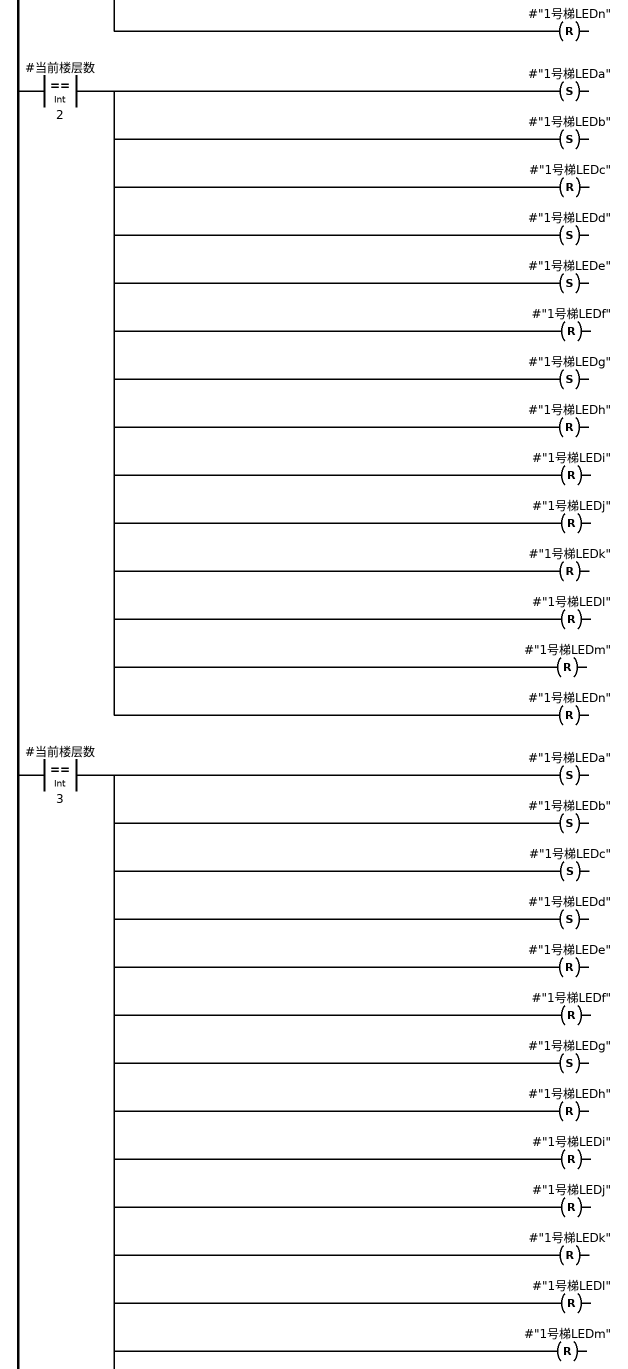
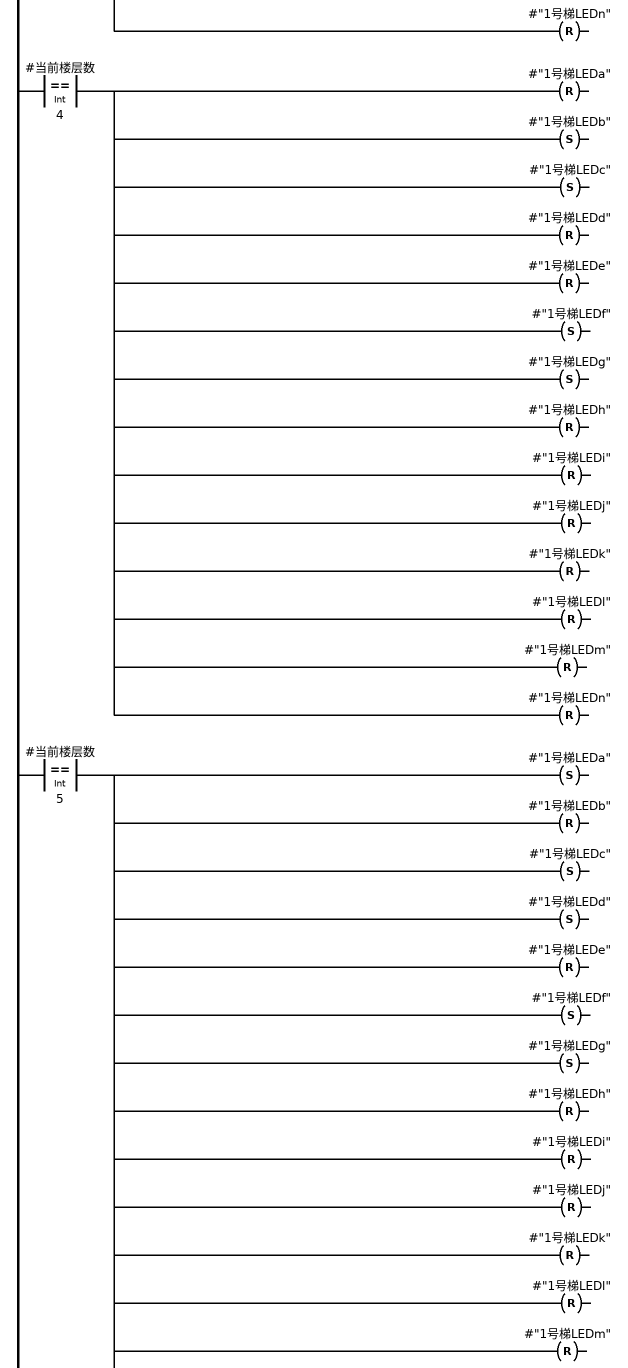
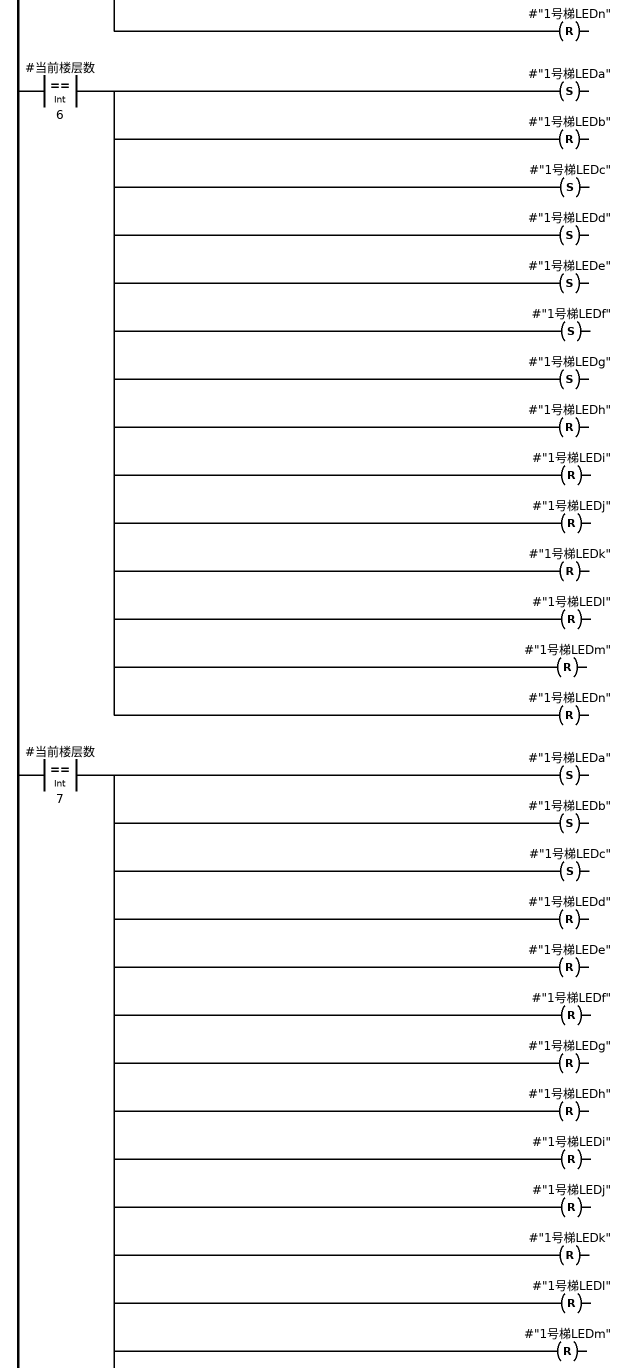
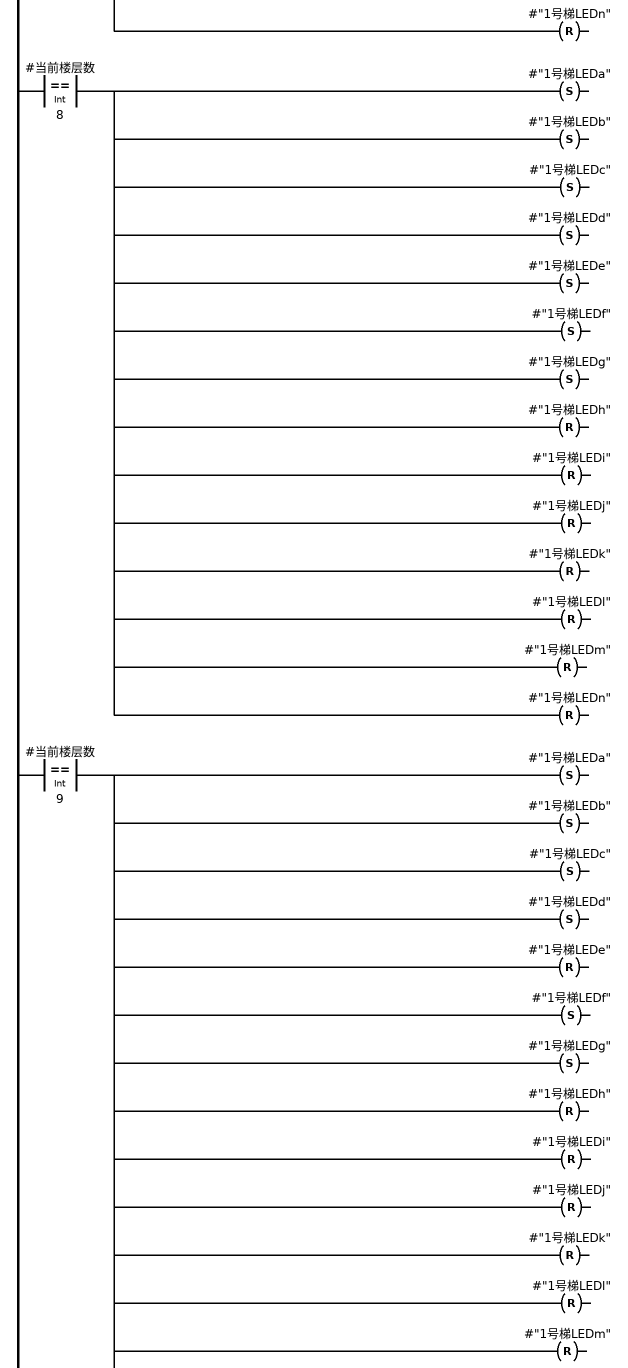
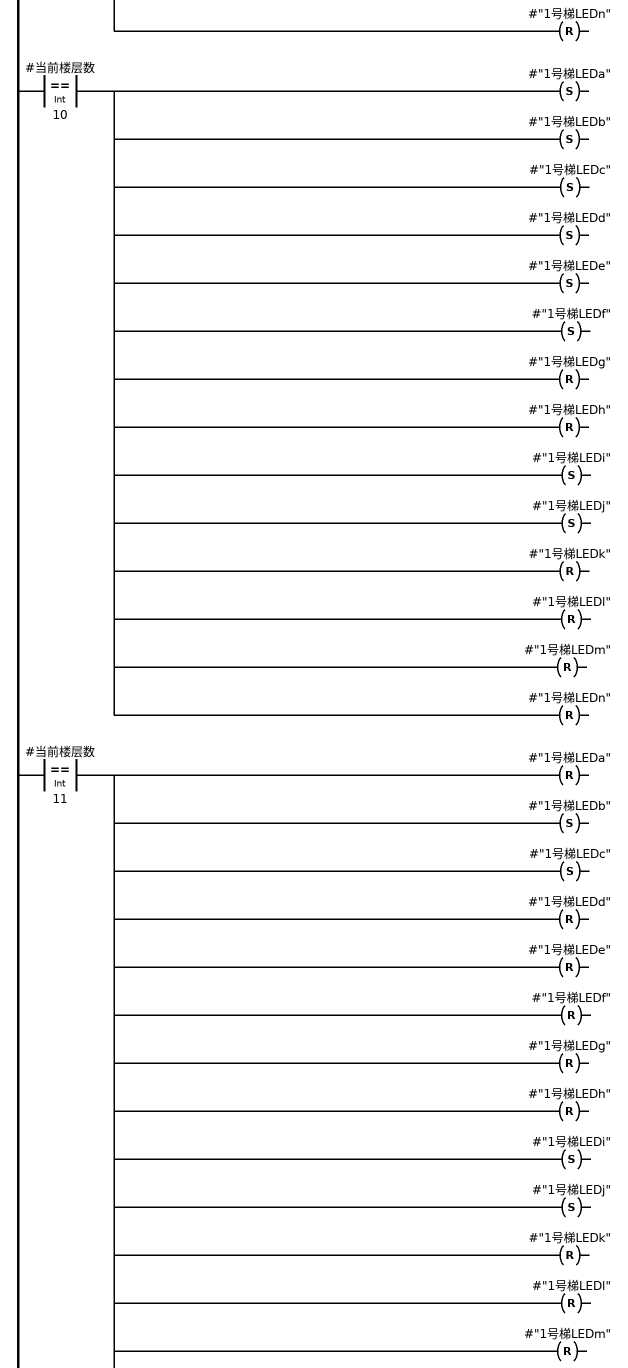
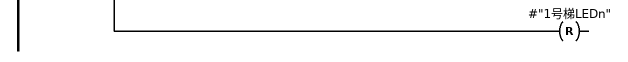
   RUNG wire#powerrail
      { S7_Templates := "SrcType := Int" } EQ_Contact(in1 := #当前楼层数, in2 := 1)
      wire#w1
      R_Coil( #"1号梯LEDa" )
   END_RUNG
   RUNG wire#w1
      S_Coil( #"1号梯LEDb" )
   END_RUNG
   RUNG wire#w1
      S_Coil( #"1号梯LEDc" )
   END_RUNG
   RUNG wire#w1
      R_Coil( #"1号梯LEDd" )
   END_RUNG
   RUNG wire#w1
      R_Coil( #"1号梯LEDe" )
   END_RUNG
   RUNG wire#w1
      R_Coil( #"1号梯LEDf" )
   END_RUNG
   RUNG wire#w1
      R_Coil( #"1号梯LEDg" )
   END_RUNG
   RUNG wire#w1
      R_Coil( #"1号梯LEDh" )
   END_RUNG
   RUNG wire#w1
      R_Coil( #"1号梯LEDi" )
   END_RUNG
   RUNG wire#w1
      R_Coil( #"1号梯LEDj" )
   END_RUNG
   RUNG wire#w1
      R_Coil( #"1号梯LEDk" )
   END_RUNG
   RUNG wire#w1
      R_Coil( #"1号梯LEDl" )
   END_RUNG
   RUNG wire#w1
      R_Coil( #"1号梯LEDm" )
   END_RUNG
   RUNG wire#w1
      R_Coil( #"1号梯LEDn" )
   END_RUNG
   RUNG wire#powerrail
      { S7_Templates := "SrcType := Int" } EQ_Contact(in1 := #当前楼层数, in2 := 0)
      wire#w2
      S_Coil( #"1号梯LEDa" )
   END_RUNG
   RUNG wire#w2
      S_Coil( #"1号梯LEDb" )
   END_RUNG
   RUNG wire#w2
      S_Coil( #"1号梯LEDc" )
   END_RUNG
   RUNG wire#w2
      S_Coil( #"1号梯LEDd" )
   END_RUNG
   RUNG wire#w2
      S_Coil( #"1号梯LEDe" )
   END_RUNG
   RUNG wire#w2
      S_Coil( #"1号梯LEDf" )
   END_RUNG
   RUNG wire#w2
      R_Coil( #"1号梯LEDg" )
   END_RUNG
   RUNG wire#w2
      R_Coil( #"1号梯LEDh" )
   END_RUNG
   RUNG wire#w2
      R_Coil( #"1号梯LEDi" )
   END_RUNG
   RUNG wire#w2
      R_Coil( #"1号梯LEDj" )
   END_RUNG
   RUNG wire#w2
      R_Coil( #"1号梯LEDk" )
   END_RUNG
   RUNG wire#w2
      R_Coil( #"1号梯LEDl" )
   END_RUNG
   RUNG wire#w2
      R_Coil( #"1号梯LEDm" )
   END_RUNG
   RUNG wire#w2
      R_Coil( #"1号梯LEDn" )
   END_RUNG
   RUNG wire#powerrail
      { S7_Templates := "SrcType := Int" } EQ_Contact(in1 := #当前楼层数, in2 := 2)
      wire#w3
      S_Coil( #"1号梯LEDa" )
   END_RUNG
   RUNG wire#w3
      S_Coil( #"1号梯LEDb" )
   END_RUNG
   RUNG wire#w3
      R_Coil( #"1号梯LEDc" )
   END_RUNG
   RUNG wire#w3
      S_Coil( #"1号梯LEDd" )
   END_RUNG
   RUNG wire#w3
      S_Coil( #"1号梯LEDe" )
   END_RUNG
   RUNG wire#w3
      R_Coil( #"1号梯LEDf" )
   END_RUNG
   RUNG wire#w3
      S_Coil( #"1号梯LEDg" )
   END_RUNG
   RUNG wire#w3
      R_Coil( #"1号梯LEDh" )
   END_RUNG
   RUNG wire#w3
      R_Coil( #"1号梯LEDi" )
   END_RUNG
   RUNG wire#w3
      R_Coil( #"1号梯LEDj" )
   END_RUNG
   RUNG wire#w3
      R_Coil( #"1号梯LEDk" )
   END_RUNG
   RUNG wire#w3
      R_Coil( #"1号梯LEDl" )
   END_RUNG
   RUNG wire#w3
      R_Coil( #"1号梯LEDm" )
   END_RUNG
   RUNG wire#w3
      R_Coil( #"1号梯LEDn" )
   END_RUNG
   RUNG wire#powerrail
      { S7_Templates := "SrcType := Int" } EQ_Contact(in1 := #当前楼层数, in2 := 3)
      wire#w4
      S_Coil( #"1号梯LEDa" )
   END_RUNG
   RUNG wire#w4
      S_Coil( #"1号梯LEDb" )
   END_RUNG
   RUNG wire#w4
      S_Coil( #"1号梯LEDc" )
   END_RUNG
   RUNG wire#w4
      S_Coil( #"1号梯LEDd" )
   END_RUNG
   RUNG wire#w4
      R_Coil( #"1号梯LEDe" )
   END_RUNG
   RUNG wire#w4
      R_Coil( #"1号梯LEDf" )
   END_RUNG
   RUNG wire#w4
      S_Coil( #"1号梯LEDg" )
   END_RUNG
   RUNG wire#w4
      R_Coil( #"1号梯LEDh" )
   END_RUNG
   RUNG wire#w4
      R_Coil( #"1号梯LEDi" )
   END_RUNG
   RUNG wire#w4
      R_Coil( #"1号梯LEDj" )
   END_RUNG
   RUNG wire#w4
      R_Coil( #"1号梯LEDk" )
   END_RUNG
   RUNG wire#w4
      R_Coil( #"1号梯LEDl" )
   END_RUNG
   RUNG wire#w4
      R_Coil( #"1号梯LEDm" )
   END_RUNG
   RUNG wire#w4
      R_Coil( #"1号梯LEDn" )
   END_RUNG
   RUNG wire#powerrail
      { S7_Templates := "SrcType := Int" } EQ_Contact(in1 := #当前楼层数, in2 := 4)
      wire#w5
      R_Coil( #"1号梯LEDa" )
   END_RUNG
   RUNG wire#w5
      S_Coil( #"1号梯LEDb" )
   END_RUNG
   RUNG wire#w5
      S_Coil( #"1号梯LEDc" )
   END_RUNG
   RUNG wire#w5
      R_Coil( #"1号梯LEDd" )
   END_RUNG
   RUNG wire#w5
      R_Coil( #"1号梯LEDe" )
   END_RUNG
   RUNG wire#w5
      S_Coil( #"1号梯LEDf" )
   END_RUNG
   RUNG wire#w5
      S_Coil( #"1号梯LEDg" )
   END_RUNG
   RUNG wire#w5
      R_Coil( #"1号梯LEDh" )
   END_RUNG
   RUNG wire#w5
      R_Coil( #"1号梯LEDi" )
   END_RUNG
   RUNG wire#w5
      R_Coil( #"1号梯LEDj" )
   END_RUNG
   RUNG wire#w5
      R_Coil( #"1号梯LEDk" )
   END_RUNG
   RUNG wire#w5
      R_Coil( #"1号梯LEDl" )
   END_RUNG
   RUNG wire#w5
      R_Coil( #"1号梯LEDm" )
   END_RUNG
   RUNG wire#w5
      R_Coil( #"1号梯LEDn" )
   END_RUNG
   RUNG wire#powerrail
      { S7_Templates := "SrcType := Int" } EQ_Contact(in1 := #当前楼层数, in2 := 5)
      wire#w6
      S_Coil( #"1号梯LEDa" )
   END_RUNG
   RUNG wire#w6
      R_Coil( #"1号梯LEDb" )
   END_RUNG
   RUNG wire#w6
      S_Coil( #"1号梯LEDc" )
   END_RUNG
   RUNG wire#w6
      S_Coil( #"1号梯LEDd" )
   END_RUNG
   RUNG wire#w6
      R_Coil( #"1号梯LEDe" )
   END_RUNG
   RUNG wire#w6
      S_Coil( #"1号梯LEDf" )
   END_RUNG
   RUNG wire#w6
      S_Coil( #"1号梯LEDg" )
   END_RUNG
   RUNG wire#w6
      R_Coil( #"1号梯LEDh" )
   END_RUNG
   RUNG wire#w6
      R_Coil( #"1号梯LEDi" )
   END_RUNG
   RUNG wire#w6
      R_Coil( #"1号梯LEDj" )
   END_RUNG
   RUNG wire#w6
      R_Coil( #"1号梯LEDk" )
   END_RUNG
   RUNG wire#w6
      R_Coil( #"1号梯LEDl" )
   END_RUNG
   RUNG wire#w6
      R_Coil( #"1号梯LEDm" )
   END_RUNG
   RUNG wire#w6
      R_Coil( #"1号梯LEDn" )
   END_RUNG
   RUNG wire#powerrail
      { S7_Templates := "SrcType := Int" } EQ_Contact(in1 := #当前楼层数, in2 := 6)
      wire#w7
      S_Coil( #"1号梯LEDa" )
   END_RUNG
   RUNG wire#w7
      R_Coil( #"1号梯LEDb" )
   END_RUNG
   RUNG wire#w7
      S_Coil( #"1号梯LEDc" )
   END_RUNG
   RUNG wire#w7
      S_Coil( #"1号梯LEDd" )
   END_RUNG
   RUNG wire#w7
      S_Coil( #"1号梯LEDe" )
   END_RUNG
   RUNG wire#w7
      S_Coil( #"1号梯LEDf" )
   END_RUNG
   RUNG wire#w7
      S_Coil( #"1号梯LEDg" )
   END_RUNG
   RUNG wire#w7
      R_Coil( #"1号梯LEDh" )
   END_RUNG
   RUNG wire#w7
      R_Coil( #"1号梯LEDi" )
   END_RUNG
   RUNG wire#w7
      R_Coil( #"1号梯LEDj" )
   END_RUNG
   RUNG wire#w7
      R_Coil( #"1号梯LEDk" )
   END_RUNG
   RUNG wire#w7
      R_Coil( #"1号梯LEDl" )
   END_RUNG
   RUNG wire#w7
      R_Coil( #"1号梯LEDm" )
   END_RUNG
   RUNG wire#w7
      R_Coil( #"1号梯LEDn" )
   END_RUNG
   RUNG wire#powerrail
      { S7_Templates := "SrcType := Int" } EQ_Contact(in1 := #当前楼层数, in2 := 7)
      wire#w8
      S_Coil( #"1号梯LEDa" )
   END_RUNG
   RUNG wire#w8
      S_Coil( #"1号梯LEDb" )
   END_RUNG
   RUNG wire#w8
      S_Coil( #"1号梯LEDc" )
   END_RUNG
   RUNG wire#w8
      R_Coil( #"1号梯LEDd" )
   END_RUNG
   RUNG wire#w8
      R_Coil( #"1号梯LEDe" )
   END_RUNG
   RUNG wire#w8
      R_Coil( #"1号梯LEDf" )
   END_RUNG
   RUNG wire#w8
      R_Coil( #"1号梯LEDg" )
   END_RUNG
   RUNG wire#w8
      R_Coil( #"1号梯LEDh" )
   END_RUNG
   RUNG wire#w8
      R_Coil( #"1号梯LEDi" )
   END_RUNG
   RUNG wire#w8
      R_Coil( #"1号梯LEDj" )
   END_RUNG
   RUNG wire#w8
      R_Coil( #"1号梯LEDk" )
   END_RUNG
   RUNG wire#w8
      R_Coil( #"1号梯LEDl" )
   END_RUNG
   RUNG wire#w8
      R_Coil( #"1号梯LEDm" )
   END_RUNG
   RUNG wire#w8
      R_Coil( #"1号梯LEDn" )
   END_RUNG
   RUNG wire#powerrail
      { S7_Templates := "SrcType := Int" } EQ_Contact(in1 := #当前楼层数, in2 := 8)
      wire#w9
      S_Coil( #"1号梯LEDa" )
   END_RUNG
   RUNG wire#w9
      S_Coil( #"1号梯LEDb" )
   END_RUNG
   RUNG wire#w9
      S_Coil( #"1号梯LEDc" )
   END_RUNG
   RUNG wire#w9
      S_Coil( #"1号梯LEDd" )
   END_RUNG
   RUNG wire#w9
      S_Coil( #"1号梯LEDe" )
   END_RUNG
   RUNG wire#w9
      S_Coil( #"1号梯LEDf" )
   END_RUNG
   RUNG wire#w9
      S_Coil( #"1号梯LEDg" )
   END_RUNG
   RUNG wire#w9
      R_Coil( #"1号梯LEDh" )
   END_RUNG
   RUNG wire#w9
      R_Coil( #"1号梯LEDi" )
   END_RUNG
   RUNG wire#w9
      R_Coil( #"1号梯LEDj" )
   END_RUNG
   RUNG wire#w9
      R_Coil( #"1号梯LEDk" )
   END_RUNG
   RUNG wire#w9
      R_Coil( #"1号梯LEDl" )
   END_RUNG
   RUNG wire#w9
      R_Coil( #"1号梯LEDm" )
   END_RUNG
   RUNG wire#w9
      R_Coil( #"1号梯LEDn" )
   END_RUNG
   RUNG wire#powerrail
      { S7_Templates := "SrcType := Int" } EQ_Contact(in1 := #当前楼层数, in2 := 9)
      wire#w10
      S_Coil( #"1号梯LEDa" )
   END_RUNG
   RUNG wire#w10
      S_Coil( #"1号梯LEDb" )
   END_RUNG
   RUNG wire#w10
      S_Coil( #"1号梯LEDc" )
   END_RUNG
   RUNG wire#w10
      S_Coil( #"1号梯LEDd" )
   END_RUNG
   RUNG wire#w10
      R_Coil( #"1号梯LEDe" )
   END_RUNG
   RUNG wire#w10
      S_Coil( #"1号梯LEDf" )
   END_RUNG
   RUNG wire#w10
      S_Coil( #"1号梯LEDg" )
   END_RUNG
   RUNG wire#w10
      R_Coil( #"1号梯LEDh" )
   END_RUNG
   RUNG wire#w10
      R_Coil( #"1号梯LEDi" )
   END_RUNG
   RUNG wire#w10
      R_Coil( #"1号梯LEDj" )
   END_RUNG
   RUNG wire#w10
      R_Coil( #"1号梯LEDk" )
   END_RUNG
   RUNG wire#w10
      R_Coil( #"1号梯LEDl" )
   END_RUNG
   RUNG wire#w10
      R_Coil( #"1号梯LEDm" )
   END_RUNG
   RUNG wire#w10
      R_Coil( #"1号梯LEDn" )
   END_RUNG
   RUNG wire#powerrail
      { S7_Templates := "SrcType := Int" } EQ_Contact(in1 := #当前楼层数, in2 := 10)
      wire#w11
      S_Coil( #"1号梯LEDa" )
   END_RUNG
   RUNG wire#w11
      S_Coil( #"1号梯LEDb" )
   END_RUNG
   RUNG wire#w11
      S_Coil( #"1号梯LEDc" )
   END_RUNG
   RUNG wire#w11
      S_Coil( #"1号梯LEDd" )
   END_RUNG
   RUNG wire#w11
      S_Coil( #"1号梯LEDe" )
   END_RUNG
   RUNG wire#w11
      S_Coil( #"1号梯LEDf" )
   END_RUNG
   RUNG wire#w11
      R_Coil( #"1号梯LEDg" )
   END_RUNG
   RUNG wire#w11
      R_Coil( #"1号梯LEDh" )
   END_RUNG
   RUNG wire#w11
      S_Coil( #"1号梯LEDi" )
   END_RUNG
   RUNG wire#w11
      S_Coil( #"1号梯LEDj" )
   END_RUNG
   RUNG wire#w11
      R_Coil( #"1号梯LEDk" )
   END_RUNG
   RUNG wire#w11
      R_Coil( #"1号梯LEDl" )
   END_RUNG
   RUNG wire#w11
      R_Coil( #"1号梯LEDm" )
   END_RUNG
   RUNG wire#w11
      R_Coil( #"1号梯LEDn" )
   END_RUNG
   RUNG wire#powerrail
      { S7_Templates := "SrcType := Int" } EQ_Contact(in1 := #当前楼层数, in2 := 11)
      wire#w12
      R_Coil( #"1号梯LEDa" )
   END_RUNG
   RUNG wire#w12
      S_Coil( #"1号梯LEDb" )
   END_RUNG
   RUNG wire#w12
      S_Coil( #"1号梯LEDc" )
   END_RUNG
   RUNG wire#w12
      R_Coil( #"1号梯LEDd" )
   END_RUNG
   RUNG wire#w12
      R_Coil( #"1号梯LEDe" )
   END_RUNG
   RUNG wire#w12
      R_Coil( #"1号梯LEDf" )
   END_RUNG
   RUNG wire#w12
      R_Coil( #"1号梯LEDg" )
   END_RUNG
   RUNG wire#w12
      R_Coil( #"1号梯LEDh" )
   END_RUNG
   RUNG wire#w12
      S_Coil( #"1号梯LEDi" )
   END_RUNG
   RUNG wire#w12
      S_Coil( #"1号梯LEDj" )
   END_RUNG
   RUNG wire#w12
      R_Coil( #"1号梯LEDk" )
   END_RUNG
   RUNG wire#w12
      R_Coil( #"1号梯LEDl" )
   END_RUNG
   RUNG wire#w12
      R_Coil( #"1号梯LEDm" )
   END_RUNG
   RUNG wire#w12
      R_Coil( #"1号梯LEDn" )
   END_RUNG
   // the same network as SCL:
   IF #当前楼层数 = 1 THEN
       #"1号梯LEDa" := FALSE;
       #"1号梯LEDb" := TRUE;
       #"1号梯LEDc" := TRUE;
       #"1号梯LEDd" := FALSE;
       #"1号梯LEDe" := FALSE;
       #"1号梯LEDf" := FALSE;
       #"1号梯LEDg" := FALSE;
       #"1号梯LEDh" := FALSE;
       #"1号梯LEDi" := FALSE;
       #"1号梯LEDj" := FALSE;
       #"1号梯LEDk" := FALSE;
       #"1号梯LEDl" := FALSE;
       #"1号梯LEDm" := FALSE;
       #"1号梯LEDn" := FALSE;
   END_IF;
   IF #当前楼层数 = 0 THEN
       #"1号梯LEDa" := TRUE;
       #"1号梯LEDb" := TRUE;
       #"1号梯LEDc" := TRUE;
       #"1号梯LEDd" := TRUE;
       #"1号梯LEDe" := TRUE;
       #"1号梯LEDf" := TRUE;
       #"1号梯LEDg" := FALSE;
       #"1号梯LEDh" := FALSE;
       #"1号梯LEDi" := FALSE;
       #"1号梯LEDj" := FALSE;
       #"1号梯LEDk" := FALSE;
       #"1号梯LEDl" := FALSE;
       #"1号梯LEDm" := FALSE;
       #"1号梯LEDn" := FALSE;
   END_IF;
   IF #当前楼层数 = 2 THEN
       #"1号梯LEDa" := TRUE;
       #"1号梯LEDb" := TRUE;
       #"1号梯LEDc" := FALSE;
       #"1号梯LEDd" := TRUE;
       #"1号梯LEDe" := TRUE;
       #"1号梯LEDf" := FALSE;
       #"1号梯LEDg" := TRUE;
       #"1号梯LEDh" := FALSE;
       #"1号梯LEDi" := FALSE;
       #"1号梯LEDj" := FALSE;
       #"1号梯LEDk" := FALSE;
       #"1号梯LEDl" := FALSE;
       #"1号梯LEDm" := FALSE;
       #"1号梯LEDn" := FALSE;
   END_IF;
   IF #当前楼层数 = 3 THEN
       #"1号梯LEDa" := TRUE;
       #"1号梯LEDb" := TRUE;
       #"1号梯LEDc" := TRUE;
       #"1号梯LEDd" := TRUE;
       #"1号梯LEDe" := FALSE;
       #"1号梯LEDf" := FALSE;
       #"1号梯LEDg" := TRUE;
       #"1号梯LEDh" := FALSE;
       #"1号梯LEDi" := FALSE;
       #"1号梯LEDj" := FALSE;
       #"1号梯LEDk" := FALSE;
       #"1号梯LEDl" := FALSE;
       #"1号梯LEDm" := FALSE;
       #"1号梯LEDn" := FALSE;
   END_IF;
   IF #当前楼层数 = 4 THEN
       #"1号梯LEDa" := FALSE;
       #"1号梯LEDb" := TRUE;
       #"1号梯LEDc" := TRUE;
       #"1号梯LEDd" := FALSE;
       #"1号梯LEDe" := FALSE;
       #"1号梯LEDf" := TRUE;
       #"1号梯LEDg" := TRUE;
       #"1号梯LEDh" := FALSE;
       #"1号梯LEDi" := FALSE;
       #"1号梯LEDj" := FALSE;
       #"1号梯LEDk" := FALSE;
       #"1号梯LEDl" := FALSE;
       #"1号梯LEDm" := FALSE;
       #"1号梯LEDn" := FALSE;
   END_IF;
   IF #当前楼层数 = 5 THEN
       #"1号梯LEDa" := TRUE;
       #"1号梯LEDb" := FALSE;
       #"1号梯LEDc" := TRUE;
       #"1号梯LEDd" := TRUE;
       #"1号梯LEDe" := FALSE;
       #"1号梯LEDf" := TRUE;
       #"1号梯LEDg" := TRUE;
       #"1号梯LEDh" := FALSE;
       #"1号梯LEDi" := FALSE;
       #"1号梯LEDj" := FALSE;
       #"1号梯LEDk" := FALSE;
       #"1号梯LEDl" := FALSE;
       #"1号梯LEDm" := FALSE;
       #"1号梯LEDn" := FALSE;
   END_IF;
   IF #当前楼层数 = 6 THEN
       #"1号梯LEDa" := TRUE;
       #"1号梯LEDb" := FALSE;
       #"1号梯LEDc" := TRUE;
       #"1号梯LEDd" := TRUE;
       #"1号梯LEDe" := TRUE;
       #"1号梯LEDf" := TRUE;
       #"1号梯LEDg" := TRUE;
       #"1号梯LEDh" := FALSE;
       #"1号梯LEDi" := FALSE;
       #"1号梯LEDj" := FALSE;
       #"1号梯LEDk" := FALSE;
       #"1号梯LEDl" := FALSE;
       #"1号梯LEDm" := FALSE;
       #"1号梯LEDn" := FALSE;
   END_IF;
   IF #当前楼层数 = 7 THEN
       #"1号梯LEDa" := TRUE;
       #"1号梯LEDb" := TRUE;
       #"1号梯LEDc" := TRUE;
       #"1号梯LEDd" := FALSE;
       #"1号梯LEDe" := FALSE;
       #"1号梯LEDf" := FALSE;
       #"1号梯LEDg" := FALSE;
       #"1号梯LEDh" := FALSE;
       #"1号梯LEDi" := FALSE;
       #"1号梯LEDj" := FALSE;
       #"1号梯LEDk" := FALSE;
       #"1号梯LEDl" := FALSE;
       #"1号梯LEDm" := FALSE;
       #"1号梯LEDn" := FALSE;
   END_IF;
   IF #当前楼层数 = 8 THEN
       #"1号梯LEDa" := TRUE;
       #"1号梯LEDb" := TRUE;
       #"1号梯LEDc" := TRUE;
       #"1号梯LEDd" := TRUE;
       #"1号梯LEDe" := TRUE;
       #"1号梯LEDf" := TRUE;
       #"1号梯LEDg" := TRUE;
       #"1号梯LEDh" := FALSE;
       #"1号梯LEDi" := FALSE;
       #"1号梯LEDj" := FALSE;
       #"1号梯LEDk" := FALSE;
       #"1号梯LEDl" := FALSE;
       #"1号梯LEDm" := FALSE;
       #"1号梯LEDn" := FALSE;
   END_IF;
   IF #当前楼层数 = 9 THEN
       #"1号梯LEDa" := TRUE;
       #"1号梯LEDb" := TRUE;
       #"1号梯LEDc" := TRUE;
       #"1号梯LEDd" := TRUE;
       #"1号梯LEDe" := FALSE;
       #"1号梯LEDf" := TRUE;
       #"1号梯LEDg" := TRUE;
       #"1号梯LEDh" := FALSE;
       #"1号梯LEDi" := FALSE;
       #"1号梯LEDj" := FALSE;
       #"1号梯LEDk" := FALSE;
       #"1号梯LEDl" := FALSE;
       #"1号梯LEDm" := FALSE;
       #"1号梯LEDn" := FALSE;
   END_IF;
   IF #当前楼层数 = 10 THEN
       #"1号梯LEDa" := TRUE;
       #"1号梯LEDb" := TRUE;
       #"1号梯LEDc" := TRUE;
       #"1号梯LEDd" := TRUE;
       #"1号梯LEDe" := TRUE;
       #"1号梯LEDf" := TRUE;
       #"1号梯LEDg" := FALSE;
       #"1号梯LEDh" := FALSE;
       #"1号梯LEDi" := TRUE;
       #"1号梯LEDj" := TRUE;
       #"1号梯LEDk" := FALSE;
       #"1号梯LEDl" := FALSE;
       #"1号梯LEDm" := FALSE;
       #"1号梯LEDn" := FALSE;
   END_IF;
   IF #当前楼层数 = 11 THEN
       #"1号梯LEDa" := FALSE;
       #"1号梯LEDb" := TRUE;
       #"1号梯LEDc" := TRUE;
       #"1号梯LEDd" := FALSE;
       #"1号梯LEDe" := FALSE;
       #"1号梯LEDf" := FALSE;
       #"1号梯LEDg" := FALSE;
       #"1号梯LEDh" := FALSE;
       #"1号梯LEDi" := TRUE;
       #"1号梯LEDj" := TRUE;
       #"1号梯LEDk" := FALSE;
       #"1号梯LEDl" := FALSE;
       #"1号梯LEDm" := FALSE;
       #"1号梯LEDn" := FALSE;
   END_IF;
END_REGION

REGION Network 3: 检修信号亮起后
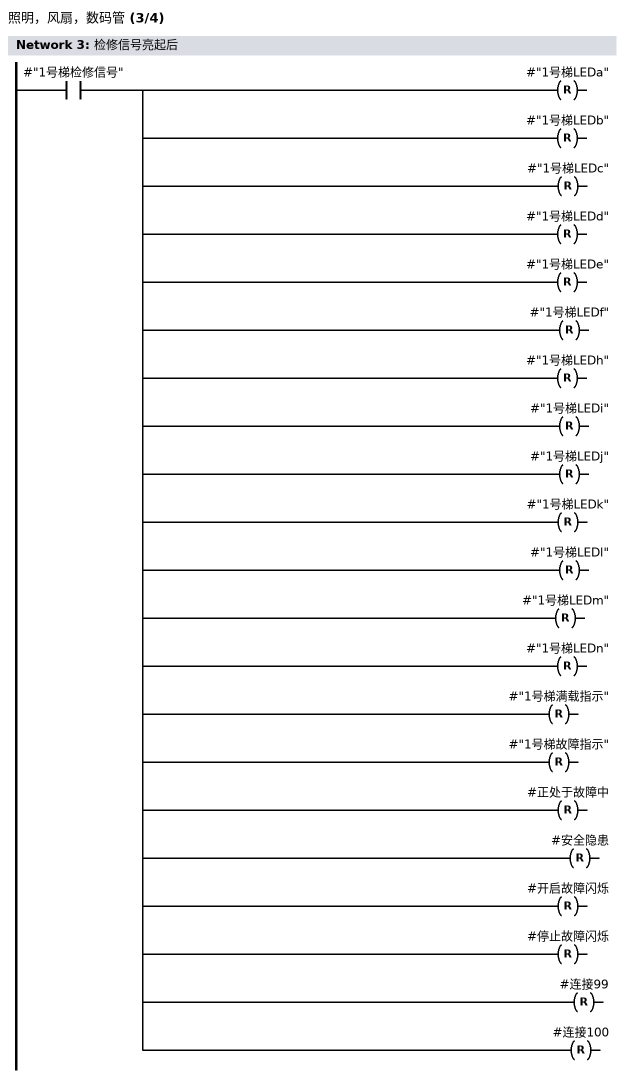
   RUNG wire#powerrail
      Contact( #"1号梯检修信号" )
      wire#w1
      R_Coil( #"1号梯LEDa" )
   END_RUNG
   RUNG wire#w1
      R_Coil( #"1号梯LEDb" )
   END_RUNG
   RUNG wire#w1
      R_Coil( #"1号梯LEDc" )
   END_RUNG
   RUNG wire#w1
      R_Coil( #"1号梯LEDd" )
   END_RUNG
   RUNG wire#w1
      R_Coil( #"1号梯LEDe" )
   END_RUNG
   RUNG wire#w1
      R_Coil( #"1号梯LEDf" )
   END_RUNG
   RUNG wire#w1
      R_Coil( #"1号梯LEDh" )
   END_RUNG
   RUNG wire#w1
      R_Coil( #"1号梯LEDi" )
   END_RUNG
   RUNG wire#w1
      R_Coil( #"1号梯LEDj" )
   END_RUNG
   RUNG wire#w1
      R_Coil( #"1号梯LEDk" )
   END_RUNG
   RUNG wire#w1
      R_Coil( #"1号梯LEDl" )
   END_RUNG
   RUNG wire#w1
      R_Coil( #"1号梯LEDm" )
   END_RUNG
   RUNG wire#w1
      R_Coil( #"1号梯LEDn" )
   END_RUNG
   RUNG wire#w1
      R_Coil( #"1号梯满载指示" )
   END_RUNG
   RUNG wire#w1
      R_Coil( #"1号梯故障指示" )
   END_RUNG
   RUNG wire#w1
      R_Coil( #正处于故障中 )
   END_RUNG
   RUNG wire#w1
      R_Coil( #安全隐患 )
   END_RUNG
   RUNG wire#w1
      R_Coil( #开启故障闪烁 )
   END_RUNG
   RUNG wire#w1
      R_Coil( #停止故障闪烁 )
   END_RUNG
   RUNG wire#w1
      R_Coil( #连接99 )
   END_RUNG
   RUNG wire#w1
      R_Coil( #连接100 )
   END_RUNG
   // the same network as SCL:
   IF #"1号梯检修信号" THEN
       #"1号梯LEDa" := FALSE;
       #"1号梯LEDb" := FALSE;
       #"1号梯LEDc" := FALSE;
       #"1号梯LEDd" := FALSE;
       #"1号梯LEDe" := FALSE;
       #"1号梯LEDf" := FALSE;
       #"1号梯LEDh" := FALSE;
       #"1号梯LEDi" := FALSE;
       #"1号梯LEDj" := FALSE;
       #"1号梯LEDk" := FALSE;
       #"1号梯LEDl" := FALSE;
       #"1号梯LEDm" := FALSE;
       #"1号梯LEDn" := FALSE;
       #"1号梯满载指示" := FALSE;
       #"1号梯故障指示" := FALSE;
       #正处于故障中 := FALSE;
       #安全隐患 := FALSE;
       #开启故障闪烁 := FALSE;
       #停止故障闪烁 := FALSE;
       #连接99 := FALSE;
       #连接100 := FALSE;
   END_IF;
END_REGION

REGION Network 4: 满载与故障
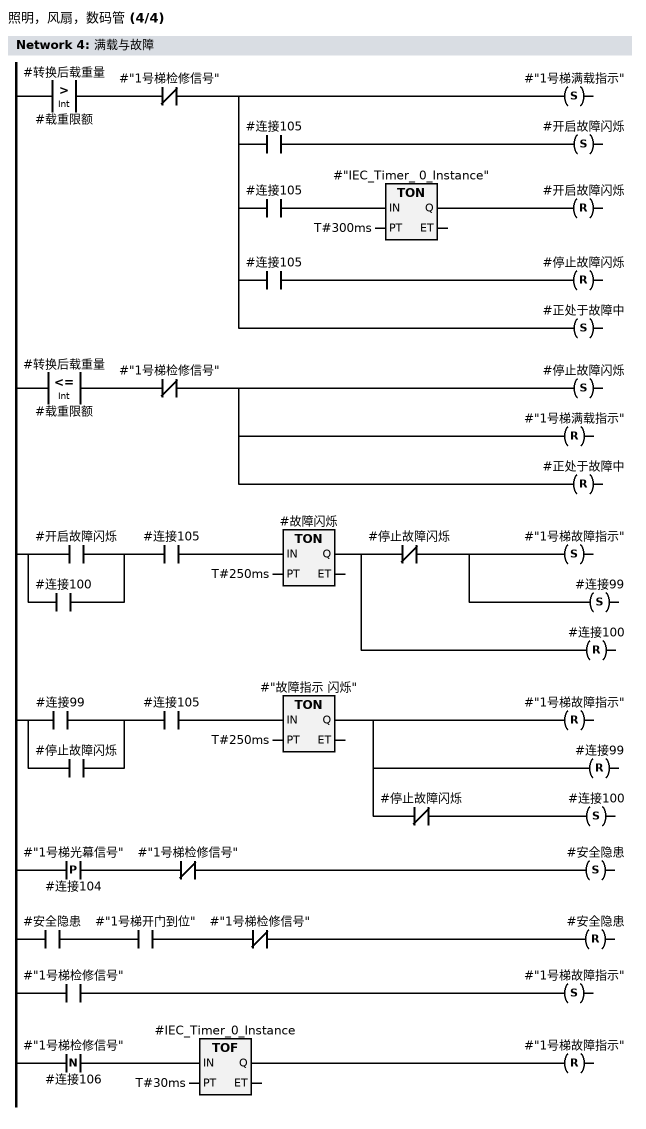
   #_w1 := (#转换后载重量 > #载重限额) AND NOT #"1号梯检修信号";
   IF #_w1 THEN #"1号梯满载指示" := TRUE; END_IF;
   IF #_w1 AND #连接105 THEN #开启故障闪烁 := TRUE; END_IF;
   #"IEC_Timer_ 0_Instance"(IN := #_w1 AND #连接105, PT := T#300ms);   // TON
   IF #"IEC_Timer_ 0_Instance".Q THEN #开启故障闪烁 := FALSE; END_IF;
   IF #_w1 AND #连接105 THEN #停止故障闪烁 := FALSE; END_IF;
   IF #_w1 THEN #正处于故障中 := TRUE; END_IF;
   IF (#转换后载重量 <= #载重限额) AND NOT #"1号梯检修信号" THEN
       #停止故障闪烁 := TRUE;
       #"1号梯满载指示" := FALSE;
       #正处于故障中 := FALSE;
   END_IF;
   #故障闪烁(IN := (#开启故障闪烁 OR #连接100) AND #连接105, PT := T#250ms);   // TON
   IF #故障闪烁.Q AND NOT #停止故障闪烁 THEN
       #"1号梯故障指示" := TRUE;
       #连接99 := TRUE;
   END_IF;
   IF #故障闪烁.Q THEN #连接100 := FALSE; END_IF;
   #"故障指示 闪烁"(IN := (#连接99 OR #停止故障闪烁) AND #连接105, PT := T#250ms);   // TON
   IF #"故障指示 闪烁".Q THEN
       #"1号梯故障指示" := FALSE;
       #连接99 := FALSE;
   END_IF;
   IF #"故障指示 闪烁".Q AND NOT #停止故障闪烁 THEN #连接100 := TRUE; END_IF;
   #_w2 := #"1号梯光幕信号" AND NOT #连接104;   // rising edge of #"1号梯光幕信号"
   #连接104 := #"1号梯光幕信号";
   IF #_w2 AND NOT #"1号梯检修信号" THEN #安全隐患 := TRUE; END_IF;
   IF #安全隐患 AND #"1号梯开门到位" AND NOT #"1号梯检修信号" THEN #安全隐患 := FALSE; END_IF;
   IF #"1号梯检修信号" THEN #"1号梯故障指示" := TRUE; END_IF;
   #_w3 := NOT #"1号梯检修信号" AND #连接106;   // falling edge of #"1号梯检修信号"
   #连接106 := #"1号梯检修信号";
   #IEC_Timer_0_Instance(IN := #_w3, PT := T#30ms);   // TOF
   IF #IEC_Timer_0_Instance.Q THEN #"1号梯故障指示" := FALSE; END_IF;
END_REGION
END_FUNCTION_BLOCK

FUNCTION_BLOCK "楼层计算"   // FB23, LAD
{ S7_Optimized_Access := 'TRUE' }
VERSION : 0.1
   VAR_INPUT
      "1号梯上平层信号" : Bool;
      "1号梯下平层信号" : Bool;
      "1号梯上端站第1限位" : Bool;
      "1号梯下端站第1限位" : Bool;
      "1号梯上行接触器" : Bool;
      "1号梯下行接触器" : Bool;
      准备就绪 : Bool;
      上端站第一限位 : Bool;
      下端站第一限位 : Bool;
      门锁1 : Bool;
      门锁2 : Bool;
      门锁3 : Bool;
      门锁4 : Bool;
      门锁5 : Bool;
      门锁6 : Bool;
      门锁7 : Bool;
      门锁8 : Bool;
      门锁9 : Bool;
      门锁10 : Bool;
   END_VAR
   VAR_OUTPUT
      上下平层同时为1 : Bool;
      当前楼层数 : Int;
      分配当前楼层数 : Int;
      正确当前楼层 : Int;
   END_VAR
   VAR RETAIN
      截下 : Bool;
   END_VAR
   VAR
      截上 : Bool;
      连接1 : Bool;
      连接2 : Bool;
      连接3 : Bool;
      连接4 : Bool;
      连接5 : Bool;
      连接6 : Bool;
      连接7 : Bool;
      连接8 : Bool;
      连接9 : Bool;
      连接10 : Bool;
      误差 : Int;
      防止不正常加数 : TOF_TIME;
      IEC_Timer_0_Instane : TON_TIME;
      "IEC_T imer_0_Instance_1" : TON_TIME;
      "IEC _Timer_0_Instance_2" : TON_TIME;
      "IEC_Timer_0 _Instance_3" : TON_TIME;
      "防止不正常减 数" : TOF_TIME;
      "IEC_Timer_ 0_Instance_5" : TON_TIME;
      "IEC_Timer_0_Instance_ 4" : TON_TIME;
      IEC_Timer_0_Instance_1 : TOF_TIME;
      IEC_Timer_0_Instance : TON_TIME;
   END_VAR
   VAR RETAIN
      计算楼层 : CTUD_INT;
   END_VAR
   VAR_TEMP   // added for the SCL form of the ladder/FBD networks
      _w1 : Bool;
      _w2 : Bool;
      _w3 : Bool;
      _w4 : Bool;
      _w5 : Bool;
      _w6 : Bool;
      _w7 : Bool;
      _w8 : Bool;
   END_VAR
BEGIN

REGION Network 1: 分配楼层
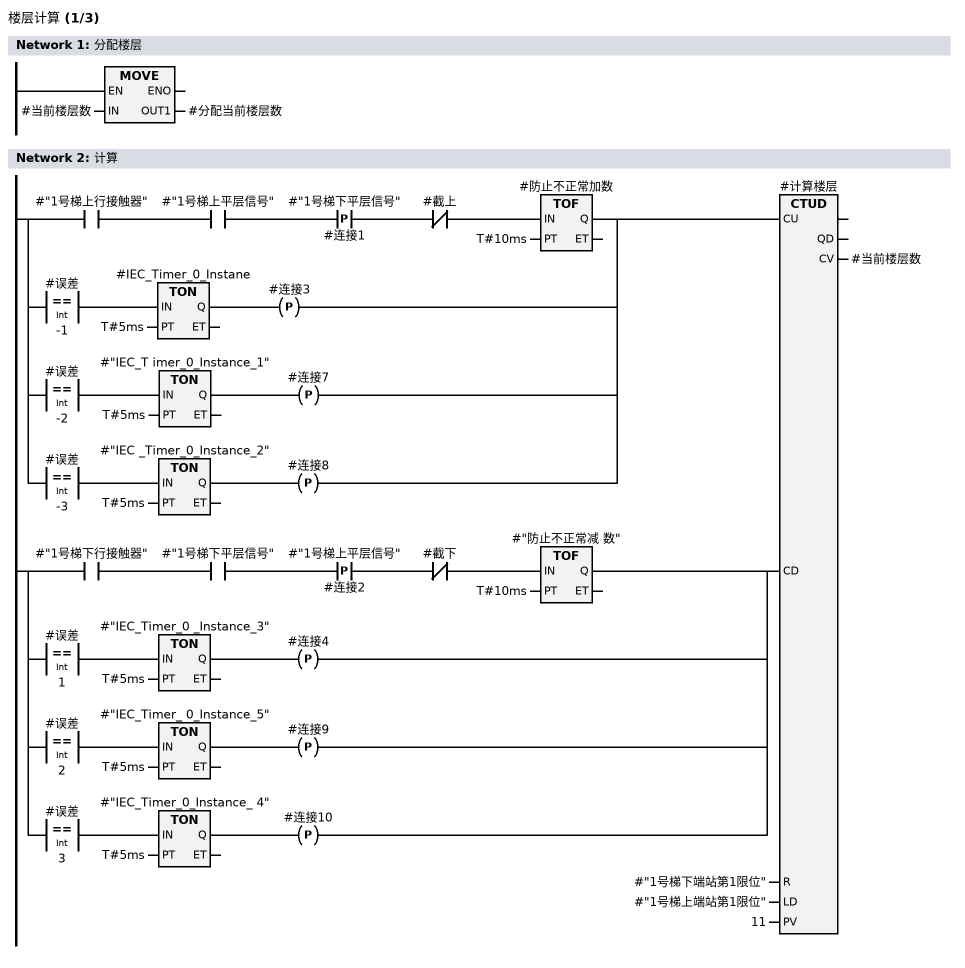
   RUNG wire#powerrail
      Move(in := #当前楼层数, out1 => #分配当前楼层数)
   END_RUNG
   // the same network as SCL:
   #分配当前楼层数 := #当前楼层数;
END_REGION

REGION Network 2: 计算
   #_w1 := #"1号梯上行接触器" AND #"1号梯上平层信号" AND #"1号梯下平层信号" AND NOT #连接1;   // rising edge of #"1号梯下平层信号"
   #连接1 := #"1号梯下平层信号";
   #防止不正常加数(IN := #_w1 AND NOT #截上, PT := T#10ms);   // TOF
   #IEC_Timer_0_Instane(IN := #误差 = (-1), PT := T#5ms);   // TON
   #_w2 := #IEC_Timer_0_Instane.Q AND NOT #连接3;   // rising edge
   #连接3 := #IEC_Timer_0_Instane.Q;
   #"IEC_T imer_0_Instance_1"(IN := #误差 = (-2), PT := T#5ms);   // TON
   #_w3 := #"IEC_T imer_0_Instance_1".Q AND NOT #连接7;   // rising edge
   #连接7 := #"IEC_T imer_0_Instance_1".Q;
   #"IEC _Timer_0_Instance_2"(IN := #误差 = (-3), PT := T#5ms);   // TON
   #_w4 := #"IEC _Timer_0_Instance_2".Q AND NOT #连接8;   // rising edge
   #连接8 := #"IEC _Timer_0_Instance_2".Q;
   #_w5 := #"1号梯下行接触器" AND #"1号梯下平层信号" AND #"1号梯上平层信号" AND NOT #连接2;   // rising edge of #"1号梯上平层信号"
   #连接2 := #"1号梯上平层信号";
   #"防止不正常减 数"(IN := #_w5 AND NOT #截下, PT := T#10ms);   // TOF
   #"IEC_Timer_0 _Instance_3"(IN := #误差 = 1, PT := T#5ms);   // TON
   #_w6 := #"IEC_Timer_0 _Instance_3".Q AND NOT #连接4;   // rising edge
   #连接4 := #"IEC_Timer_0 _Instance_3".Q;
   #"IEC_Timer_ 0_Instance_5"(IN := #误差 = 2, PT := T#5ms);   // TON
   #_w7 := #"IEC_Timer_ 0_Instance_5".Q AND NOT #连接9;   // rising edge
   #连接9 := #"IEC_Timer_ 0_Instance_5".Q;
   #"IEC_Timer_0_Instance_ 4"(IN := #误差 = 3, PT := T#5ms);   // TON
   #_w8 := #"IEC_Timer_0_Instance_ 4".Q AND NOT #连接10;   // rising edge
   #连接10 := #"IEC_Timer_0_Instance_ 4".Q;
   #计算楼层(CU := #防止不正常加数.Q OR #_w2 OR #_w3 OR #_w4,   // CTUD
         CD := #"防止不正常减 数".Q OR #_w6 OR #_w7 OR #_w8,
         R := #"1号梯下端站第1限位",
         LD := #"1号梯上端站第1限位",
         PV := 11,
         CV => #当前楼层数);
END_REGION

REGION Network 3: 截上截下
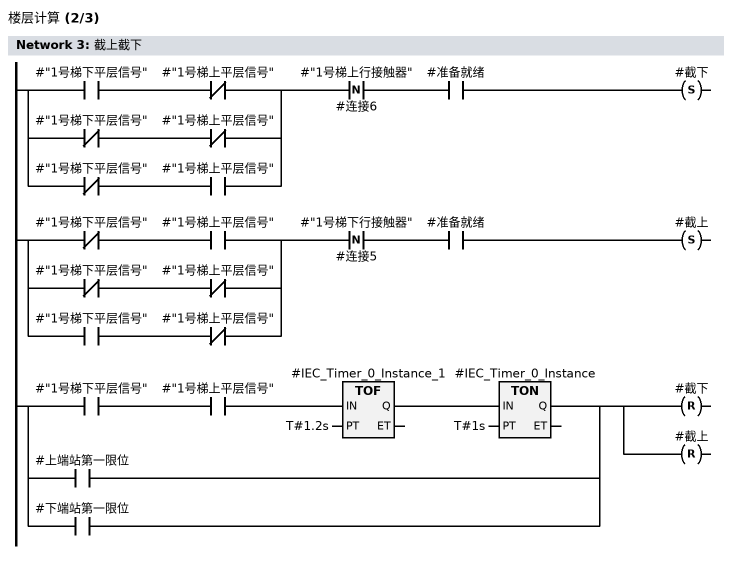
   #_w1 := ((#"1号梯下平层信号" AND NOT #"1号梯上平层信号") OR (NOT #"1号梯下平层信号" AND NOT #"1号梯上平层信号") OR (NOT #"1号梯下平层信号" AND #"1号梯上平层信号")) AND NOT #"1号梯上行接触器" AND #连接6;   // falling edge of #"1号梯上行接触器"
   #连接6 := #"1号梯上行接触器";
   IF #_w1 AND #准备就绪 THEN #截下 := TRUE; END_IF;
   #_w2 := ((NOT #"1号梯下平层信号" AND #"1号梯上平层信号") OR (NOT #"1号梯下平层信号" AND NOT #"1号梯上平层信号") OR (#"1号梯下平层信号" AND NOT #"1号梯上平层信号")) AND NOT #"1号梯下行接触器" AND #连接5;   // falling edge of #"1号梯下行接触器"
   #连接5 := #"1号梯下行接触器";
   IF #_w2 AND #准备就绪 THEN #截上 := TRUE; END_IF;
   #IEC_Timer_0_Instance_1(IN := #"1号梯下平层信号" AND #"1号梯上平层信号", PT := T#1.2s);   // TOF
   #IEC_Timer_0_Instance(IN := #IEC_Timer_0_Instance_1.Q, PT := T#1s);   // TON
   IF #IEC_Timer_0_Instance.Q OR #上端站第一限位 OR #下端站第一限位 THEN
       #截下 := FALSE;
       #截上 := FALSE;
   END_IF;
END_REGION

REGION Network 4: 判断楼层，纠正
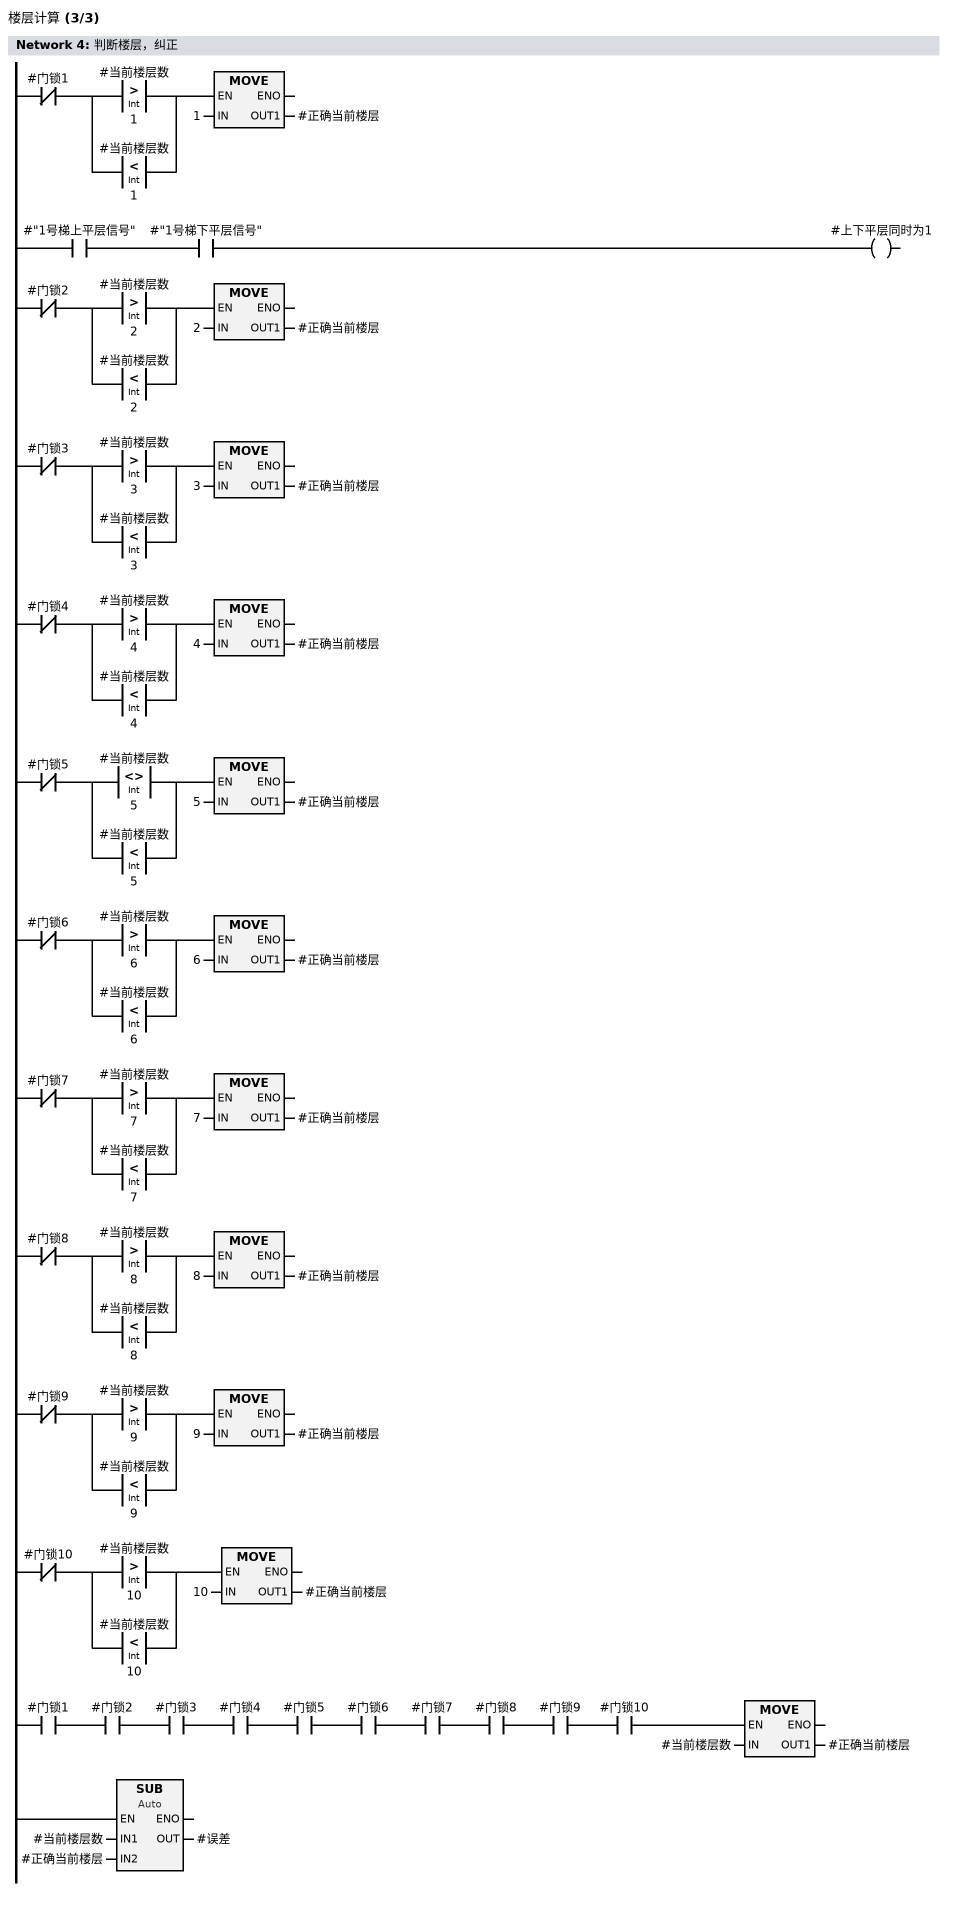
   RUNG wire#powerrail
      I_Contact( #门锁1 )
      wire#w1
      { S7_Templates := "SrcType := Int" } GT_Contact(in1 := #当前楼层数, in2 := 1)
      wire#w2
      Move(in := 1, out1 => #正确当前楼层)
   END_RUNG
   RUNG wire#w1
      { S7_Templates := "SrcType := Int" } LT_Contact(in1 := #当前楼层数, in2 := 1)
   END_RUNG wire#w2
   RUNG wire#powerrail
      Contact( #"1号梯上平层信号" )
      Contact( #"1号梯下平层信号" )
      Coil( #上下平层同时为1 )
   END_RUNG
   RUNG wire#powerrail
      I_Contact( #门锁2 )
      wire#w3
      { S7_Templates := "SrcType := Int" } GT_Contact(in1 := #当前楼层数, in2 := 2)
      wire#w4
      Move(in := 2, out1 => #正确当前楼层)
   END_RUNG
   RUNG wire#w3
      { S7_Templates := "SrcType := Int" } LT_Contact(in1 := #当前楼层数, in2 := 2)
   END_RUNG wire#w4
   RUNG wire#powerrail
      I_Contact( #门锁3 )
      wire#w5
      { S7_Templates := "SrcType := Int" } GT_Contact(in1 := #当前楼层数, in2 := 3)
      wire#w6
      Move(in := 3, out1 => #正确当前楼层)
   END_RUNG
   RUNG wire#w5
      { S7_Templates := "SrcType := Int" } LT_Contact(in1 := #当前楼层数, in2 := 3)
   END_RUNG wire#w6
   RUNG wire#powerrail
      I_Contact( #门锁4 )
      wire#w7
      { S7_Templates := "SrcType := Int" } GT_Contact(in1 := #当前楼层数, in2 := 4)
      wire#w8
      Move(in := 4, out1 => #正确当前楼层)
   END_RUNG
   RUNG wire#w7
      { S7_Templates := "SrcType := Int" } LT_Contact(in1 := #当前楼层数, in2 := 4)
   END_RUNG wire#w8
   RUNG wire#powerrail
      I_Contact( #门锁5 )
      wire#w9
      { S7_Templates := "SrcType := Int" } NE_Contact(in1 := #当前楼层数, in2 := 5)
      wire#w10
      Move(in := 5, out1 => #正确当前楼层)
   END_RUNG
   RUNG wire#w9
      { S7_Templates := "SrcType := Int" } LT_Contact(in1 := #当前楼层数, in2 := 5)
   END_RUNG wire#w10
   RUNG wire#powerrail
      I_Contact( #门锁6 )
      wire#w11
      { S7_Templates := "SrcType := Int" } GT_Contact(in1 := #当前楼层数, in2 := 6)
      wire#w12
      Move(in := 6, out1 => #正确当前楼层)
   END_RUNG
   RUNG wire#w11
      { S7_Templates := "SrcType := Int" } LT_Contact(in1 := #当前楼层数, in2 := 6)
   END_RUNG wire#w12
   RUNG wire#powerrail
      I_Contact( #门锁7 )
      wire#w13
      { S7_Templates := "SrcType := Int" } GT_Contact(in1 := #当前楼层数, in2 := 7)
      wire#w14
      Move(in := 7, out1 => #正确当前楼层)
   END_RUNG
   RUNG wire#w13
      { S7_Templates := "SrcType := Int" } LT_Contact(in1 := #当前楼层数, in2 := 7)
   END_RUNG wire#w14
   RUNG wire#powerrail
      I_Contact( #门锁8 )
      wire#w15
      { S7_Templates := "SrcType := Int" } GT_Contact(in1 := #当前楼层数, in2 := 8)
      wire#w16
      Move(in := 8, out1 => #正确当前楼层)
   END_RUNG
   RUNG wire#w15
      { S7_Templates := "SrcType := Int" } LT_Contact(in1 := #当前楼层数, in2 := 8)
   END_RUNG wire#w16
   RUNG wire#powerrail
      I_Contact( #门锁9 )
      wire#w17
      { S7_Templates := "SrcType := Int" } GT_Contact(in1 := #当前楼层数, in2 := 9)
      wire#w18
      Move(in := 9, out1 => #正确当前楼层)
   END_RUNG
   RUNG wire#w17
      { S7_Templates := "SrcType := Int" } LT_Contact(in1 := #当前楼层数, in2 := 9)
   END_RUNG wire#w18
   RUNG wire#powerrail
      I_Contact( #门锁10 )
      wire#w19
      { S7_Templates := "SrcType := Int" } GT_Contact(in1 := #当前楼层数, in2 := 10)
      wire#w20
      Move(in := 10, out1 => #正确当前楼层)
   END_RUNG
   RUNG wire#w19
      { S7_Templates := "SrcType := Int" } LT_Contact(in1 := #当前楼层数, in2 := 10)
   END_RUNG wire#w20
   RUNG wire#powerrail
      Contact( #门锁1 )
      Contact( #门锁2 )
      Contact( #门锁3 )
      Contact( #门锁4 )
      Contact( #门锁5 )
      Contact( #门锁6 )
      Contact( #门锁7 )
      Contact( #门锁8 )
      Contact( #门锁9 )
      Contact( #门锁10 )
      Move(in := #当前楼层数, out1 => #正确当前楼层)
   END_RUNG
   RUNG wire#powerrail
      Sub(in1 := #当前楼层数, in2 := #正确当前楼层, out => #误差)
   END_RUNG
   // the same network as SCL:
   IF NOT #门锁1 AND ((#当前楼层数 > 1) OR (#当前楼层数 < 1)) THEN #正确当前楼层 := 1; END_IF;
   #上下平层同时为1 := #"1号梯上平层信号" AND #"1号梯下平层信号";
   IF NOT #门锁2 AND ((#当前楼层数 > 2) OR (#当前楼层数 < 2)) THEN #正确当前楼层 := 2; END_IF;
   IF NOT #门锁3 AND ((#当前楼层数 > 3) OR (#当前楼层数 < 3)) THEN #正确当前楼层 := 3; END_IF;
   IF NOT #门锁4 AND ((#当前楼层数 > 4) OR (#当前楼层数 < 4)) THEN #正确当前楼层 := 4; END_IF;
   IF NOT #门锁5 AND ((#当前楼层数 <> 5) OR (#当前楼层数 < 5)) THEN #正确当前楼层 := 5; END_IF;
   IF NOT #门锁6 AND ((#当前楼层数 > 6) OR (#当前楼层数 < 6)) THEN #正确当前楼层 := 6; END_IF;
   IF NOT #门锁7 AND ((#当前楼层数 > 7) OR (#当前楼层数 < 7)) THEN #正确当前楼层 := 7; END_IF;
   IF NOT #门锁8 AND ((#当前楼层数 > 8) OR (#当前楼层数 < 8)) THEN #正确当前楼层 := 8; END_IF;
   IF NOT #门锁9 AND ((#当前楼层数 > 9) OR (#当前楼层数 < 9)) THEN #正确当前楼层 := 9; END_IF;
   IF NOT #门锁10 AND ((#当前楼层数 > 10) OR (#当前楼层数 < 10)) THEN #正确当前楼层 := 10; END_IF;
   IF #门锁1 AND #门锁2 AND #门锁3 AND #门锁4 AND #门锁5 AND #门锁6 AND #门锁7 AND #门锁8 AND #门锁9 AND #门锁10 THEN
       #正确当前楼层 := #当前楼层数;
   END_IF;
   #误差 := #当前楼层数 - #正确当前楼层;
END_REGION
END_FUNCTION_BLOCK

FUNCTION_BLOCK "距离调度"   // FB27, LAD
{ S7_Optimized_Access := 'TRUE' }
VERSION : 0.1
   VAR_INPUT
      准备就绪 : Bool;
      检修信号 : Bool;
      上下平层都为1 : Bool;
      上呼灯1 : Bool;
      上呼灯2 : Bool;
      上呼灯3 : Bool;
      上呼灯4 : Bool;
      上呼灯5 : Bool;
      上呼灯6 : Bool;
      上呼灯7 : Bool;
      上呼灯8 : Bool;
      上呼灯9 : Bool;
      下呼灯2 : Bool;
      下呼灯3 : Bool;
      下呼灯4 : Bool;
      下呼灯5 : Bool;
      下呼灯6 : Bool;
      下呼灯7 : Bool;
      下呼灯8 : Bool;
      下呼灯9 : Bool;
      下呼灯10 : Bool;
      上行指示 : Bool;
      下行指示 : Bool;
      当前楼层 : Int;
      外呼上面有目标最大数1 : Int;
      外呼上面有目标最大数2 : Int;
      外呼上面有目标最大数3 : Int;
      外呼上面有目标最大数4 : Int;
      外呼上面有目标最大数5 : Int;
      外呼上面有目标最大数6 : Int;
      外呼上面有目标最大数7 : Int;
      外呼上面有目标最大数8 : Int;
      外呼上面有目标最大数9 : Int;
      外呼下面有目标最小数2 : Int;
      外呼下面有目标最小数3 : Int;
      外呼下面有目标最小数4 : Int;
      外呼下面有目标最小数5 : Int;
      外呼下面有目标最小数6 : Int;
      外呼下面有目标最小数7 : Int;
      外呼下面有目标最小数8 : Int;
      外呼下面有目标最小数9 : Int;
      外呼下面有目标最小数10 : Int;
      外呼下面有目标2 : Bool;
      外呼下面有目标3 : Bool;
      外呼下面有目标4 : Bool;
      外呼下面有目标5 : Bool;
      外呼下面有目标6 : Bool;
      外呼下面有目标7 : Bool;
      外呼下面有目标8 : Bool;
      外呼下面有目标9 : Bool;
      外呼下面有目标10 : Bool;
      外呼上面有目标1 : Bool;
      外呼上面有目标2 : Bool;
      外呼上面有目标3 : Bool;
      外呼上面有目标4 : Bool;
      外呼上面有目标5 : Bool;
      外呼上面有目标6 : Bool;
      外呼上面有目标7 : Bool;
      外呼上面有目标8 : Bool;
      外呼上面有目标9 : Bool;
      外呼下面无目标2 : Bool;
      外呼下面无目标3 : Bool;
      外呼下面无目标4 : Bool;
      外呼下面无目标5 : Bool;
      外呼下面无目标6 : Bool;
      外呼下面无目标7 : Bool;
      外呼下面无目标8 : Bool;
      外呼下面无目标9 : Bool;
      外呼上面无目标2 : Bool;
      外呼上面无目标3 : Bool;
      外呼上面无目标4 : Bool;
      外呼上面无目标5 : Bool;
      外呼上面无目标6 : Bool;
      外呼上面无目标7 : Bool;
      外呼上面无目标8 : Bool;
      外呼上面无目标9 : Bool;
      上行停站次数3 : Int;
      上行停站次数4 : Int;
      上行停站次数5 : Int;
      上行停站次数6 : Int;
      上行停站次数7 : Int;
      上行停站次数8 : Int;
      上行停站次数9 : Int;
      下行停站次数2 : Int;
      下行停站次数3 : Int;
      下行停站次数4 : Int;
      下行停站次数5 : Int;
      下行停站次数6 : Int;
      下行停站次数7 : Int;
      下行停站次数8 : Int;
      上行停站次数10 : Int;
      下行停站次数1 : Int;
      载重量 : Int;
      死机 : Bool;
      限重分配 : Int;
   END_VAR
   VAR_OUTPUT
      最终调度距离上1 : Int;
      最终调度距离上2 : Int;
      最终调度距离上3 : Int;
      最终调度距离上4 : Int;
      最终调度距离上5 : Int;
      最终调度距离上6 : Int;
      最终调度距离上7 : Int;
      最终调度距离上8 : Int;
      最终调度距离上9 : Int;
      最终调度距离下2 : Int;
      最终调度距离下3 : Int;
      最终调度距离下4 : Int;
      最终调度距离下5 : Int;
      最终调度距离下6 : Int;
      最终调度距离下7 : Int;
      最终调度距离下8 : Int;
      最终调度距离下9 : Int;
      最终调度距离下10 : Int;
   END_VAR
   VAR
      检修中 : Bool;
      "2层边沿触发1" : Bool;
      "2层边沿触发2" : Bool;
      "2层边沿触发3" : Bool;
      "2层边沿触发4" : Bool;
      "2层边沿触发5" : Bool;
      "2层边沿触发6" : Bool;
      "2层边沿触发7" : Bool;
      "2层边沿触发8" : Bool;
      "2层边沿触发9" : Bool;
      "2层边沿触发10" : Bool;
      "2层调度距离1" : Int;
      "2层调度距离2" : Int;
      "2层调度距离3" : Int;
      "2层调度距离4" : Int;
      "2层调度距离5" : Int;
      "2层调度距离6" : Int;
      "2层调度距离7" : Int;
      "2层调度距离8" : Int;
      "2层调度距离9" : Int;
      "2层调度距离10" : Int;
      "3层边沿触发1" : Bool;
      "3层边沿触发2" : Bool;
      "3层边沿触发3" : Bool;
      "3层边沿触发4" : Bool;
      "3层边沿触发5" : Bool;
      "3层边沿触发6" : Bool;
      "3层边沿触发7" : Bool;
      "3层边沿触发8" : Bool;
      "3层边沿触发9" : Bool;
      "3层边沿触发10" : Bool;
      "3层调度距离1" : Int;
      "3层调度距离2" : Int;
      "3层调度距离3" : Int;
      "3层调度距离4" : Int;
      "3层调度距离5" : Int;
      "3层调度距离6" : Int;
      "3层调度距离7" : Int;
      "3层调度距离8" : Int;
      "3层调度距离9" : Int;
      "3层调度距离10" : Int;
      "4层边沿触发1" : Bool;
      "4层边沿触发2" : Bool;
      "4层边沿触发3" : Bool;
      "4层边沿触发4" : Bool;
      "4层边沿触发5" : Bool;
      "4层边沿触发6" : Bool;
      "4层边沿触发7" : Bool;
      "4层边沿触发8" : Bool;
      "4层边沿触发9" : Bool;
      "4层边沿触发10" : Bool;
      "4层调度距离1" : Int;
      "4层调度距离2" : Int;
      "4层调度距离3" : Int;
      "4层调度距离4" : Int;
      "4层调度距离5" : Int;
      "4层调度距离6" : Int;
      "4层调度距离7" : Int;
      "4层调度距离8" : Int;
      "4层调度距离9" : Int;
      "4层调度距离10" : Int;
      "5层调度距离1" : Int;
      "5层调度距离2" : Int;
      "5层调度距离3" : Int;
      "5层调度距离4" : Int;
      "5层调度距离5" : Int;
      "5层调度距离6" : Int;
      "5层调度距离7" : Int;
      "5层调度距离8" : Int;
      "5层调度距离9" : Int;
      "5层调度距离10" : Int;
      "5层边沿触发1" : Bool;
      "5层边沿触发2" : Bool;
      "5层边沿触发3" : Bool;
      "5层边沿触发4" : Bool;
      "5层边沿触发5" : Bool;
      "5层边沿触发6" : Bool;
      "5层边沿触发7" : Bool;
      "5层边沿触发8" : Bool;
      "5层边沿触发9" : Bool;
      "5层边沿触发10" : Bool;
      "6层边沿触发1" : Bool;
      "6层边沿触发2" : Bool;
      "6层边沿触发3" : Bool;
      "6层边沿触发4" : Bool;
      "6层边沿触发5" : Bool;
      "6层边沿触发6" : Bool;
      "6层边沿触发7" : Bool;
      "6层边沿触发8" : Bool;
      "6层边沿触发9" : Bool;
      "6层边沿触发10" : Bool;
      "6层调度距离1" : Int;
      "6层调度距离2" : Int;
      "6层调度距离3" : Int;
      "6层调度距离4" : Int;
      "6层调度距离5" : Int;
      "6层调度距离6" : Int;
      "6层调度距离7" : Int;
      "6层调度距离8" : Int;
      "6层调度距离9" : Int;
      "6层调度距离10" : Int;
      "7层调度距离1" : Int;
      "7层调度距离2" : Int;
      "7层调度距离3" : Int;
      "7层调度距离4" : Int;
      "7层调度距离5" : Int;
      "7层调度距离6" : Int;
      "7层调度距离7" : Int;
      "7层调度距离8" : Int;
      "7层调度距离9" : Int;
      "7层调度距离10" : Int;
      "7层边沿触发1" : Bool;
      "7层边沿触发2" : Bool;
      "7层边沿触发3" : Bool;
      "7层边沿触发4" : Bool;
      "7层边沿触发5" : Bool;
      "7层边沿触发6" : Bool;
      "7层边沿触发7" : Bool;
      "7层边沿触发8" : Bool;
      "7层边沿触发9" : Bool;
      "7层边沿触发10" : Bool;
      "8层边沿触发1" : Bool;
      "8层边沿触发2" : Bool;
      "8层边沿触发3" : Bool;
      "8层边沿触发4" : Bool;
      "8层边沿触发5" : Bool;
      "8层边沿触发6" : Bool;
      "8层边沿触发7" : Bool;
      "8层边沿触发8" : Bool;
      "8层边沿触发9" : Bool;
      "8层边沿触发10" : Bool;
      "8层调度距离1" : Int;
      "8层调度距离2" : Int;
      "8层调度距离3" : Int;
      "8层调度距离4" : Int;
      "8层调度距离5" : Int;
      "8层调度距离6" : Int;
      "8层调度距离7" : Int;
      "8层调度距离8" : Int;
      "8层调度距离9" : Int;
      "8层调度距离10" : Int;
      "9层调度距离1" : Int;
      "9层调度距离2" : Int;
      "9层调度距离3" : Int;
      "9层调度距离4" : Int;
      "9层调度距离5" : Int;
      "9层调度距离6" : Int;
      "9层调度距离7" : Int;
      "9层调度距离8" : Int;
      "9层调度距离9" : Int;
      "9层调度距离10" : Int;
      "9层边沿触发1" : Bool;
      "9层边沿触发2" : Bool;
      "9层边沿触发3" : Bool;
      "9层边沿触发4" : Bool;
      "9层边沿触发5" : Bool;
      "9层边沿触发6" : Bool;
      "9层边沿触发7" : Bool;
      "9层边沿触发8" : Bool;
      "9层边沿触发9" : Bool;
      "9层边沿触发10" : Bool;
      "1层调度距离1" : Int;
      "1层调度距离2" : Int;
      "1层边沿触发1" : Bool;
      "1层边沿触发2" : Bool;
      "10层边沿触发1" : Bool;
      "10层边沿触发2" : Bool;
      "10层调度距离1" : Int;
      "10层调度距离2" : Int;
   END_VAR
   VAR_TEMP   // added for the SCL form of the ladder/FBD networks
      _w1 : Bool;
      _w2 : Bool;
      _w3 : Bool;
      _w4 : Bool;
      _w5 : Bool;
      _w6 : Bool;
      _w7 : Bool;
      _w8 : Bool;
      _w9 : Bool;
      _w10 : Bool;
      _w11 : Bool;
      _w12 : Bool;
   END_VAR
BEGIN

REGION Network 1: 2层调度距离
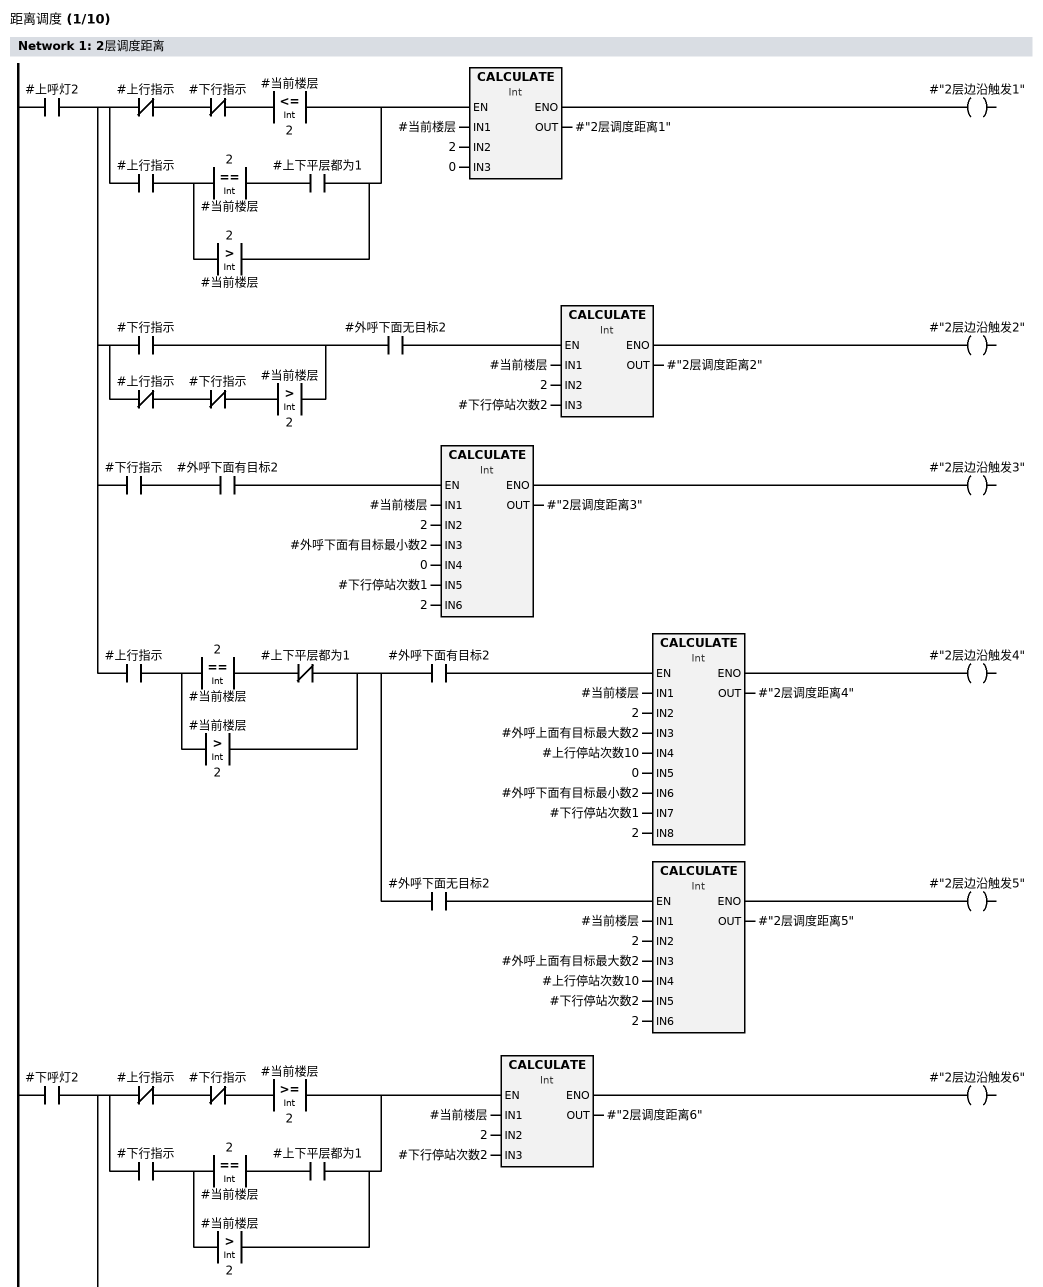
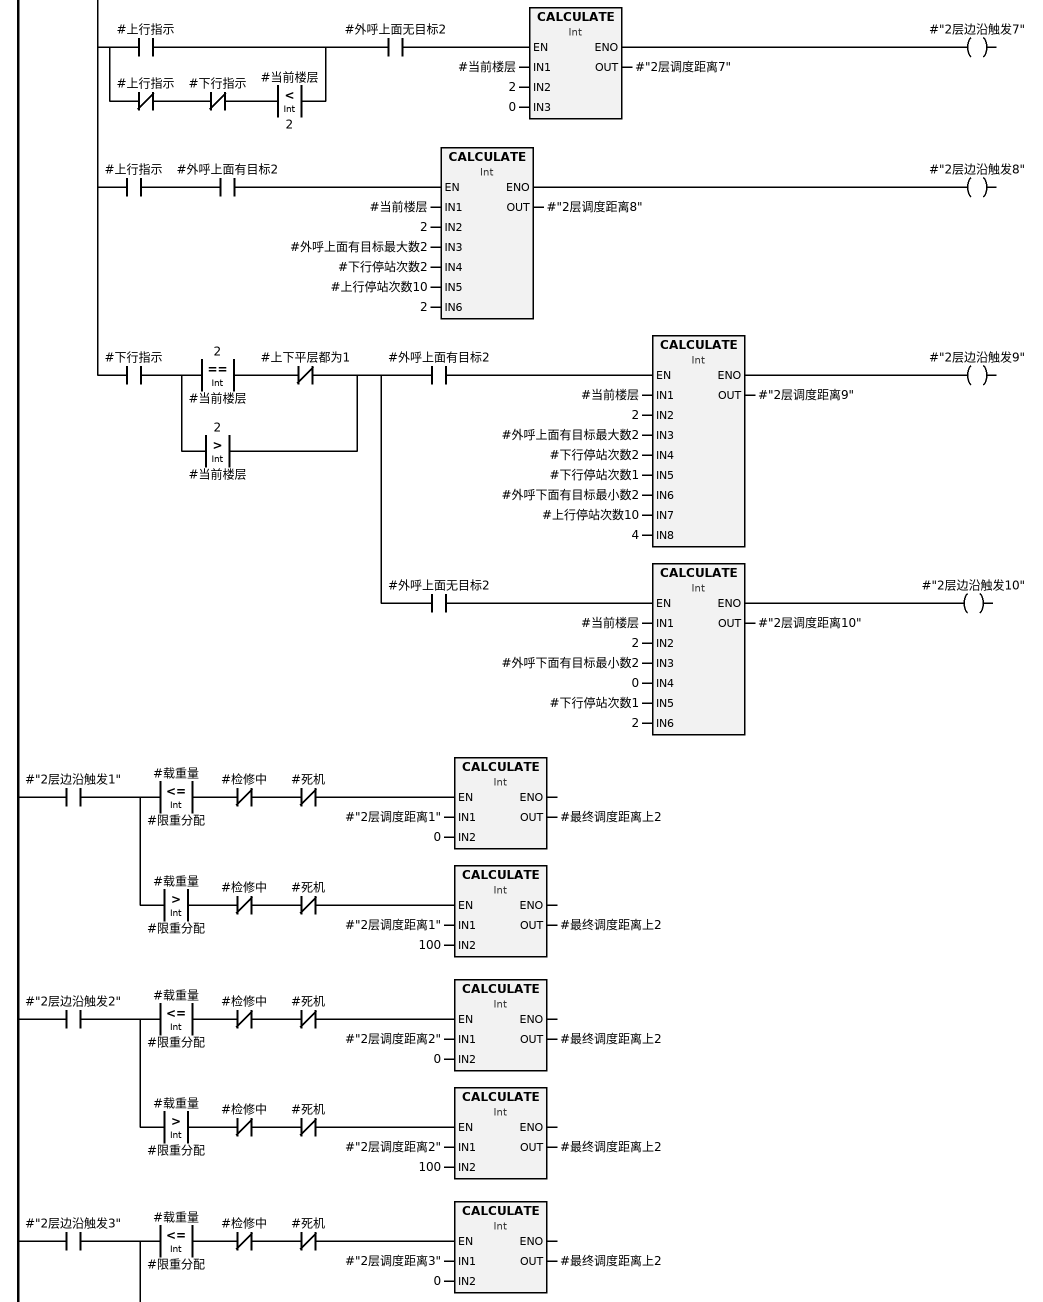
